(* IEC 61131-3 sources: daoli-st-library/DL_Process (part 22) *)

(* ---- FB_DL_BatteryTestCycler.st ---- *)
//==============================================================================
// 功能块：FB_DL_BatteryTestCycler ｜ 中文名称：单通道电池充放电工步机
// 所属子库：DL_Process ｜ 版本：v1.0.1 ｜ 兼容：CODESYS V3.5+ / TwinCAT 3 / 汇川 InoProShop
// 功能描述：单体电芯充放电测试工步机：静置 → 恒流充电 → 恒压充电 → 静置 → 恒流放电 →
//           静置 → 完成，逐工步按终止判据切相；充/放电容量按安时积分统计（LREAL 累加
//           防精度损失）；温度与电压安全域逐拍硬判，越限当拍断流并进故障相（锂电热失控
//           不可逆，安全路径优先级最高）。工步超时按「本工步独立计时」判定，禁跨相累计。
//           本件是单通道工步机：不调度多通道、不做通道仲裁与分配（多通道调度归
//           序号 19 的 FormationsChannelMgr），对外只以电流设定 / 电压限值与工步状态
//           布尔快照交互，两件互不包含。
// 开源溯源 (Origin)：道莅原创实现（参考 公开工程惯例 分类与参数域）
// 单位表：电压[V] / 电流[A]（放电为负）/ 温度[摄氏度] / 静置时长[min] / 工步超时[min] /
//         容量[Ah] / 容量比[百分数] / 扫描间隔[ms] / 工步已历时[ms] / 样本数[拍]
// 错误码表：16#0005_0406 信息级（工步切相提示，含「因终止判据达成而提前切相」与静置
//           到时，不置 bError）/ 16#0005_0407 信息级（容量统计饱和触顶，不置 bError）/
//           16#0005_034B 故障级（温度越上限或电压越安全域，或安全判据量（温度/电压/
//           电流）非有限——非有限按越限处置，强制断流，置 bError）/ 16#0005_034C 故障级
//           （单工步超时，工艺卡死，置 bError + 断流）/ 16#0005_034D 故障级（组态非法：
//           额定容量/电流设定/电压域/超时非正或非有限，以及状态机 ELSE 非法状态兜底）。
//           034D 的共用反证句：组态非法与非法状态在现有输出组合下不可观测出差异（均为
//           bError + fCurrentSetA = 0 + eStep 不推进 + bValid 撤），§3 未给本件独立组态槽，
//           故显式复用不越段。
// 状态机：E_DL_BatteryCycleState（eIdle=0 待机 / eRestInit=10 充电前静置 / eCcCharge=20
//           恒流充电 / eCvCharge=30 恒压充电 / eRestMid=40 放前静置 / eDiscCharge=50 恒流
//           放电 / eRestFinal=60 放后静置 / eDone=70 完成 / eFault=99 故障兜底），CASE 含
//           ELSE 兜底，ELSE 置 034D 且断流、eStep 回 eIdle。
// 边界行为：① 安全侧优先：温度 > fTempMaxC 或电压越 [fVoltMinV, fVoltMaxV] → 故障 034B
//           + fCurrentSetA := 0.0 + 进 eFault（每拍先判安全判据，先于任何工步推进）；
//           ② 单工步超 tMaxStep → 故障 034C，工步计时器在每次切相时清零（禁相内累计，
//           R40 家族）；③ 额定容量/电流/电压域/超时组态非法 → 034D 组态分支（映射见
//           错误码表反证句）；④ 容量积分 Ah += |I| x Δt/3600，LREAL 累加并饱和；⑤ CV
//           终止：|I| < fCutoffCurrentA 连续 nCvHoldSamples 拍才切相（防单点抖动误切）；
//           ⑥ bStop → 当拍 fCurrentSetA := 0 并回 eIdle（不等待工步收尾）；⑦ 失能走同一
//           安全侧路径（fCurrentSetA := 0）。bStart 取上升沿，bStepDone 为单拍脉冲。
// 修订历史：v1.0.0 2026-11-17 首版（R25 派单 · §4.15）
//           v1.0.1 2026-11-17 终审补 eFault 独立 CASE 标签（对外引脚契约零变更）：原实现 eFault(99)
//           无标签，落进 ELSE 兜底支路每拍把真因码 034B/034C 覆盖成 034D「非法状态」，激励消失后
//           诊断失真（故障仍锁存、安全侧不变，属诊断保真度缺陷）。同批另有 6 件存在同类标签缺失
//           （ParticleCounterStat / CoolingTowerApproachCalc / InverterGridSync / HeatPumpDefrost /
//           DuctStaticReset / DewpointReset），已按 R106 第二档挂账下轮统一修并加机检规则。
//==============================================================================
(*------------------------------------------------------------------------------
 * 枚举: E_DL_BatteryCycleState（归属 DL_Process，与 FB_DL_BatteryTestCycler 同文件）
 *       工步号与 §4.15 顺序一一对应；数值步长留空位便于插工步
 *----------------------------------------------------------------------------*)
TYPE E_DL_BatteryCycleState :
(
    eIdle       := 0,   // 待机：电流设定 0，等待 bStart / Idle, current setpoint 0, waiting for start
    eRestInit   := 10,  // 充电前静置：时长 tRestCharge / Pre-charge rest, duration tRestCharge
    eCcCharge   := 20,  // 恒流充电：电流 = fCcCurrentA，终止判据 电压达 fCvVoltV / Constant-current charge
    eCvCharge   := 30,  // 恒压充电：电压限 = fCvVoltV，终止判据 电流降至 fCutoffCurrentA / Constant-voltage charge
    eRestMid    := 40,  // 放前静置：时长 tRestCharge / Pre-discharge rest, duration tRestCharge
    eDiscCharge := 50,  // 恒流放电：电流 = -fDiscCurrentA，终止判据 电压降至 fDiscCutoffV / Constant-current discharge
    eRestFinal  := 60,  // 放后静置：时长 tRestDisc / Post-discharge rest, duration tRestDisc
    eDone       := 70,  // 完成：电流设定 0，容量统计保持 / Done, current 0, capacity statistics held
    eFault      := 99   // 故障兜底：越限/超时/组态非法/非法状态 / Fault fallback
);
END_TYPE

(*==============================================================================
 * 功能块: FB_DL_BatteryTestCycler
 * 调用约定: 每个扫描周期无条件调用一次；uDeltaTimeMs 必须注入真实任务间隔。
 *============================================================================*)
FUNCTION_BLOCK FB_DL_BatteryTestCycler
VAR_INPUT
    fVoltV          : LREAL;                       // 实测电压 [V] / Measured voltage [V]
    fCurrentA       : LREAL;                       // 实测电流 [A]，放电为负 / Measured current [A], negative while discharging
    fTempC          : LREAL;                       // 实测温度 [摄氏度] / Measured temperature [degC]
    fCcCurrentA     : LREAL;                       // 恒流充电电流设定 [A]，须 > 0 / Constant-current charge setpoint [A], must be > 0
    fCvVoltV        : LREAL;                       // 恒压充电电压点 [V] / Constant-voltage charge point [V]
    fCutoffCurrentA : LREAL;                       // 恒压段终止电流 [A]，须 >= 0 / CV termination current [A], must be >= 0
    fDiscCurrentA   : LREAL;                       // 放电电流设定 [A]，须 > 0（本件按负值下发）/ Discharge current setpoint [A], must be > 0, issued negative
    fDiscCutoffV    : LREAL;                       // 放电终止电压 [V] / Discharge termination voltage [V]
    tRestCharge     : TIME := T#10M;               // 充/放前静置时长 [min] / Pre-step rest duration [min]
    tRestDisc       : TIME := T#10M;               // 放后静置时长 [min] / Post-discharge rest duration [min]
    tMaxStep        : TIME := T#120M;              // 单工步超时 [min]，各工步独立计时 / Per-step timeout [min], timed per step
    fCapNomAh       : LREAL;                       // 额定容量 [Ah]，须 > 0（容量比分母）/ Rated capacity [Ah], must be > 0
    fVoltMaxV       : LREAL;                       // 安全域电压上限 [V] / Safety voltage ceiling [V]
    fVoltMinV       : LREAL;                       // 安全域电压下限 [V] / Safety voltage floor [V]
    fTempMaxC       : LREAL;                       // 温度上限 [摄氏度] / Temperature ceiling [degC]
    bStart          : BOOL;                        // 启动（取上升沿）/ Start, rising edge
    bStop           : BOOL;                        // 停止（电平，当拍断流）/ Stop, level, current dropped this scan
    bReset          : BOOL;                        // 复位，上升沿清故障与容量统计 / Reset, rising edge clears the fault and capacity statistics
    uDeltaTimeMs    : UDINT;                       // 扫描间隔 [ms]，调用方注入，禁系统时间函数 / Scan interval [ms], caller-injected
END_VAR
VAR_OUTPUT
    eStep           : E_DL_BatteryCycleState;      // 当前工步 / Current step
    fCurrentSetA    : LREAL;                       // 电流设定 [A]，故障拍立即 0 / Current setpoint [A], forced to 0 on any fault scan
    fVoltLimitV     : LREAL;                       // 电压限 [V]，随工步切换 / Voltage limit [V], follows the step
    fChargedAh      : LREAL;                       // 累计充电容量 [Ah]，饱和 / Accumulated charge capacity [Ah], saturating
    fDischargedAh   : LREAL;                       // 累计放电容量 [Ah]，饱和 / Accumulated discharge capacity [Ah], saturating
    fCapacityRatioPct : LREAL;                     // 容量比 [百分数] = 放电 Ah / 额定 Ah x 100 / Capacity ratio [percent]
    bStepDone       : BOOL;                        // 工步完成单拍脉冲（切相当拍 TRUE）/ Single-scan step-done pulse
    tStepElapsed    : TIME;                        // 本工步已历时 [ms] / Elapsed time of the current step [ms]
    eErr            : UDINT;                       // 错误码，0 = 无错，码位 16#0005_0406 起信息级、16#0005_034B 起故障级（分带见错误码表） / Error code, 0 = no error, band info/fault per the code table
    bError          : BOOL;                        // 故障级标志，仅故障级错误置位 / Fault-class flag, set only on fault-level codes
    bValid          : BOOL;                        // 工步输出可用标志，失能/故障闸显式 FALSE / Step outputs usable flag, explicit FALSE on disable/fault gates
END_VAR
VAR
    fbReset         : R_TRIG;                      // 复位上升沿检测实例 / Reset rising edge detector
    fbStart         : R_TRIG;                      // 启动上升沿检测实例 / Start rising edge detector
    uStepMs         : UDINT;                       // 本工步累计历时 [ms]，切相即清零 / Elapsed time of this step [ms], cleared on every transition
    uDtEff          : UDINT;                       // 钳位后的扫描间隔 [ms] / Clamped scan interval [ms]
    uMaxStepMs      : UDINT;                       // 工步超时门限 [ms] / Step timeout threshold [ms]
    uRestChgMs      : UDINT;                       // 充/放前静置门限 [ms] / Pre-step rest threshold [ms]
    uRestDiscMs     : UDINT;                       // 放后静置门限 [ms] / Post-discharge rest threshold [ms]
    fDtH            : LREAL;                       // 扫描间隔换算成小时 [h] / Scan interval in hours [h]
    fAbsCurrentA    : LREAL;                       // 实测电流绝对值 [A] / Absolute measured current [A]
    fAhStep         : LREAL;                       // 本拍容量增量 [Ah] / Capacity increment of this scan [Ah]
    nCvHoldCnt      : INT;                         // CV 终止判据连续满足拍数 [拍] / Consecutive CV-cutoff samples [scans]
    bCapSat         : BOOL;                        // 容量积分饱和标志 / Capacity saturation flag
    bStepChanged    : BOOL;                        // 本拍发生切相标志 / Step changed this scan
    bRestChgDone    : BOOL;                        // 静置到时（用充电侧时长）/ Rest elapsed with the charge-side duration
    bRestDiscDone   : BOOL;                        // 静置到时（用放电侧时长）/ Rest elapsed with the discharge-side duration
    bCvCutoff       : BOOL;                        // CV 终止判据满足 / CV termination criterion satisfied
    bDiscCutoff     : BOOL;                        // 放电终止判据满足 / Discharge termination criterion satisfied
    bCcReached      : BOOL;                        // CC 段电压已达 CV 点 / CC reached the CV point
    bNonFinSafe     : BOOL;                        // 安全判据量非有限标志 / Safety-class non-finite flag
    bNonFinCfg      : BOOL;                        // 组态量非有限标志 / Configuration non-finite flag
    bFirstScan      : BOOL := TRUE;                // 上电首拍标志 / First-scan flag
END_VAR
VAR CONSTANT
    DL_BTC_CODE_INFO_1 : UDINT := 16#0005_0406;    // 信息级槽 1（工步切相提示） / info slot 1
    DL_BTC_CODE_INFO_2 : UDINT := 16#0005_0407;    // 信息级槽 2（容量统计饱和） / info slot 2
    DL_BTC_CODE_FLT_1  : UDINT := 16#0005_034B;    // 故障级槽 1（温度/电压越限，强制断流） / fault slot 1
    DL_BTC_CODE_FLT_2  : UDINT := 16#0005_034C;    // 故障级槽 2（工步超时，工艺卡死） / fault slot 2
    DL_BTC_CODE_FLT_3  : UDINT := 16#0005_034D;    // 故障级槽 3（组态非法/非法状态兜底） / fault slot 3
    DL_BTC_CV_HOLD     : INT := 5;                 // CV 终止判据连续确认拍数 [拍] / CV cutoff confirmation samples [scans]
    DL_BTC_AH_MAX      : LREAL := 100000.0;        // 容量积分饱和上限 [Ah] / Capacity saturation ceiling [Ah]
    DL_BTC_DT_MIN_MS   : UDINT := 1;               // 扫描间隔下限 [ms]，防除零与死判 / Scan interval floor [ms]
    DL_BTC_SEC_PER_H   : LREAL := 3600.0;          // 秒转小时系数 [s/h] / Seconds per hour
    DL_BTC_MS_PER_S    : LREAL := 1000.0;          // 毫秒转秒系数 [ms/s] / Milliseconds per second
    DL_BTC_PCT         : LREAL := 100.0;           // 百分数系数 [百分数] / Percent factor
    DL_BTC_ZERO        : LREAL := 0.0;             // 零值常量，避免裸字面量 [—] / Zero constant, avoids a bare literal
    DL_BTC_TOL         : LREAL := 1.0E-6;          // 浮点比较容差 [—] / Float comparison tolerance
    DL_BTC_INF         : LREAL := 1.7976931348623157E308; // LREAL 幅值上限，Inf 判据 / LREAL magnitude ceiling
END_VAR

(*------------------------------------------------------------------------------
 * 段 1｜无条件刷新区（红线 5）：复位/启动沿检测在任何分支之外周期调用；
 *       bStepDone 为单拍脉冲，逐拍先清（调用方读到的仍是本拍值）
 *----------------------------------------------------------------------------*)
bStepDone := FALSE;                                // 单拍脉冲先清（自清机制）/ single-scan pulse cleared first
fCurrentSetA := DL_BTC_ZERO;                       // 电流设定默认 0：任何未显式赋值的路径都断流 / default 0, any unassigned path is de-energised
fVoltLimitV := DL_BTC_ZERO;                        // 电压限默认 0 / voltage limit defaults to zero
fbReset(CLK := bReset);                            // 复位沿检测无条件刷新 / reset edge refreshed unconditionally
fbStart(CLK := bStart);                            // 启动沿检测无条件刷新 / start edge refreshed unconditionally

(*------------------------------------------------------------------------------
 * 段 2｜复位沿处理（改写置于沿后，防吞沿 R39）：清故障与容量统计
 *----------------------------------------------------------------------------*)
IF fbReset.Q THEN
    eStep := E_DL_BatteryCycleState.eIdle;
    eErr   := 16#0000_0000;                        // 复位清码 / reset clears the code
    bError := FALSE;                               // 复位清故障 / reset clears the fault
    fChargedAh := DL_BTC_ZERO;                     // 充电容量清 / charge capacity cleared
    fDischargedAh := DL_BTC_ZERO;                  // 放电容量清 / discharge capacity cleared
    fCapacityRatioPct := DL_BTC_ZERO;              // 容量比清 / capacity ratio cleared
    uStepMs := 16#0000_0000;                       // 工步计时清 / step timer cleared
    nCvHoldCnt := 0;                               // CV 确认计数清 / CV hold counter cleared
    bCapSat := FALSE;                              // 饱和标志清 / saturation flag cleared
    bFirstScan := TRUE;                            // 重新首拍化 / re-initialize first scan
END_IF

(*------------------------------------------------------------------------------
 * 段 3｜非有限输入闸：安全判据量（温度/电压/电流）非有限 → 按越限处置（034B，断流）；
 *       组态量非有限 → 034D 组态分支。分两类是因为前者的正确处置是「当拍断流」，
 *       后者是「拒绝启动」
 *----------------------------------------------------------------------------*)
bNonFinSafe := (fVoltV <> fVoltV) OR (ABS(fVoltV) >= DL_BTC_INF)
            OR (fCurrentA <> fCurrentA) OR (ABS(fCurrentA) >= DL_BTC_INF)
            OR (fTempC <> fTempC) OR (ABS(fTempC) >= DL_BTC_INF);   // 安全判据量非有限 / safety-class non-finite
bNonFinCfg := (fCcCurrentA <> fCcCurrentA) OR (ABS(fCcCurrentA) >= DL_BTC_INF)
           OR (fCvVoltV <> fCvVoltV) OR (ABS(fCvVoltV) >= DL_BTC_INF)
           OR (fCutoffCurrentA <> fCutoffCurrentA) OR (ABS(fCutoffCurrentA) >= DL_BTC_INF)
           OR (fDiscCurrentA <> fDiscCurrentA) OR (ABS(fDiscCurrentA) >= DL_BTC_INF)
           OR (fDiscCutoffV <> fDiscCutoffV) OR (ABS(fDiscCutoffV) >= DL_BTC_INF)
           OR (fCapNomAh <> fCapNomAh) OR (ABS(fCapNomAh) >= DL_BTC_INF)
           OR (fVoltMaxV <> fVoltMaxV) OR (ABS(fVoltMaxV) >= DL_BTC_INF)
           OR (fVoltMinV <> fVoltMinV) OR (ABS(fVoltMinV) >= DL_BTC_INF)
           OR (fTempMaxC <> fTempMaxC) OR (ABS(fTempMaxC) >= DL_BTC_INF);   // 组态量非有限 / configuration non-finite
IF bNonFinSafe THEN
    eStep := E_DL_BatteryCycleState.eFault;        // 进故障相 / enter fault state
    eErr   := DL_BTC_CODE_FLT_1;                   // 故障级：安全判据不可判，按越限处置 / fault: safety values undecidable, treated as out of range
    bError := TRUE;                                // 故障级必置 bError（R45 配对）/ fault-class pairs with bError
    fCurrentSetA := DL_BTC_ZERO;                   // 当拍断流（安全路径最高优先）/ current dropped this scan
    fVoltLimitV := DL_BTC_ZERO;                    // 电压限撤 / voltage limit dropped
    bValid := FALSE;                               // 故障闸显式不可用（R72）/ explicit FALSE on the fault gate
    RETURN;
END_IF
IF bNonFinCfg THEN
    eStep := E_DL_BatteryCycleState.eFault;        // 进故障相 / enter fault state
    eErr   := DL_BTC_CODE_FLT_3;                   // 故障级：组态非法（映射见错误码表）/ fault: invalid configuration, mapping per the code table
    bError := TRUE;                                // 故障级必置 bError（R45 配对）/ fault-class pairs with bError
    fCurrentSetA := DL_BTC_ZERO;                   // 断流 / current dropped
    fVoltLimitV := DL_BTC_ZERO;                    // 电压限撤 / voltage limit dropped
    bValid := FALSE;                               // 故障闸显式不可用（R72）/ explicit FALSE on the fault gate
    RETURN;
END_IF

(*------------------------------------------------------------------------------
 * 段 4｜组态域闸（034D 组态分支，先判后除：容量比分母在此被证明为正）
 *----------------------------------------------------------------------------*)
IF (fCapNomAh <= DL_BTC_TOL) OR (fVoltMaxV <= fVoltMinV + DL_BTC_TOL)
   OR (fCcCurrentA <= DL_BTC_TOL) OR (fDiscCurrentA <= DL_BTC_TOL)
   OR (fCutoffCurrentA < DL_BTC_ZERO)
   OR (DINT_TO_UDINT(TIME_TO_DINT(tMaxStep)) = 16#00000000) THEN
    eStep := E_DL_BatteryCycleState.eFault;        // 进故障相 / enter fault state
    eErr   := DL_BTC_CODE_FLT_3;                   // 故障级：组态非法 / fault: invalid configuration
    bError := TRUE;                                // 故障级必置 bError（R45 配对）/ fault-class pairs with bError
    fCurrentSetA := DL_BTC_ZERO;                   // 断流 / current dropped
    fVoltLimitV := DL_BTC_ZERO;                    // 电压限撤 / voltage limit dropped
    bValid := FALSE;                               // 故障闸显式不可用（R72）/ explicit FALSE on the fault gate
    RETURN;
END_IF

(*------------------------------------------------------------------------------
 * 段 5｜安全域硬判（最高优先，先于任何工步推进）：温度越上限或电压越安全域 →
 *       034B + 当拍断流 + 进故障相。故障锁存至 bReset（热失控不可逆）
 *----------------------------------------------------------------------------*)
IF (fTempC > fTempMaxC) OR (fVoltV > fVoltMaxV + DL_BTC_TOL) OR (fVoltV < fVoltMinV - DL_BTC_TOL) THEN
    eStep := E_DL_BatteryCycleState.eFault;        // 进故障相 / enter fault state
    eErr   := DL_BTC_CODE_FLT_1;                   // 故障级：温度/电压越限 / fault: temperature or voltage out of range
    bError := TRUE;                                // 故障级必置 bError（R45 配对）/ fault-class pairs with bError
    fCurrentSetA := DL_BTC_ZERO;                   // 当拍断流（安全侧）/ current dropped this scan, safe side
    fVoltLimitV := DL_BTC_ZERO;                    // 电压限撤 / voltage limit dropped
    bValid := FALSE;                               // 故障闸显式不可用（R72）/ explicit FALSE on the fault gate
    RETURN;
END_IF

(*------------------------------------------------------------------------------
 * 段 6｜工步计时：仅活动工步累计（切相清零），静置/完成/待机不累计
 *----------------------------------------------------------------------------*)
IF uDeltaTimeMs < DL_BTC_DT_MIN_MS THEN
    uDtEff := DL_BTC_DT_MIN_MS;                     // 间隔过小按下限，防死等 / floored interval prevents a dead wait
ELSE
    uDtEff := uDeltaTimeMs;                         // 间隔原值 / interval as-is
END_IF
IF (eStep <> E_DL_BatteryCycleState.eIdle) AND (eStep <> E_DL_BatteryCycleState.eDone)
   AND (eStep <> E_DL_BatteryCycleState.eFault) THEN
    IF uStepMs < 16#FFFF_FFFE THEN
        uStepMs := uStepMs + uDtEff;                // 本工步累计 [ms] / accumulate the current step [ms]
    END_IF
END_IF
uMaxStepMs := DINT_TO_UDINT(TIME_TO_DINT(tMaxStep));       // 超时门限 [ms] / timeout threshold [ms]
uRestChgMs := DINT_TO_UDINT(TIME_TO_DINT(tRestCharge));    // 充/放前静置门限 [ms] / pre-step rest threshold [ms]
uRestDiscMs := DINT_TO_UDINT(TIME_TO_DINT(tRestDisc));     // 放后静置门限 [ms] / post-discharge rest threshold [ms]

(*------------------------------------------------------------------------------
 * 段 7｜工步超时（034C）：各工步独立计时，切相即清零，禁相内累计（R40 家族）
 *----------------------------------------------------------------------------*)
IF (eStep <> E_DL_BatteryCycleState.eIdle) AND (eStep <> E_DL_BatteryCycleState.eDone)
   AND (eStep <> E_DL_BatteryCycleState.eFault) AND (uStepMs > uMaxStepMs) THEN
    eStep := E_DL_BatteryCycleState.eFault;        // 进故障相 / enter fault state
    eErr   := DL_BTC_CODE_FLT_2;                   // 故障级：工步超时，工艺卡死 / fault: step timeout, process stuck
    bError := TRUE;                                // 故障级必置 bError（R45 配对）/ fault-class pairs with bError
    fCurrentSetA := DL_BTC_ZERO;                   // 断流 / current dropped
    fVoltLimitV := DL_BTC_ZERO;                    // 电压限撤 / voltage limit dropped
    bValid := FALSE;                               // 故障闸显式不可用（R72）/ explicit FALSE on the fault gate
    RETURN;
END_IF

(*------------------------------------------------------------------------------
 * 段 8｜容量安时积分：Ah += |I| x Δt/3600（LREAL 累加防精度损失，饱和防溢出）
 *----------------------------------------------------------------------------*)
fDtH := UDINT_TO_LREAL(uDtEff) / DL_BTC_MS_PER_S / DL_BTC_SEC_PER_H;   // 间隔换算成小时 [h] / interval in hours
fAbsCurrentA := ABS(fCurrentA);                    // 电流绝对值 [A] / absolute current [A]
fAhStep := fAbsCurrentA * fDtH;                     // 本拍容量增量 [Ah] / capacity increment [Ah]
IF (eStep = E_DL_BatteryCycleState.eCcCharge) OR (eStep = E_DL_BatteryCycleState.eCvCharge) THEN
    IF fChargedAh < DL_BTC_AH_MAX THEN
        fChargedAh := fChargedAh + fAhStep;         // 充电容量累加 [Ah] / charge capacity accumulation
        IF fChargedAh >= DL_BTC_AH_MAX THEN
            fChargedAh := DL_BTC_AH_MAX;            // 饱和钳位 [Ah] / saturation clamp
            bCapSat := TRUE;                        // 饱和标志 / saturation flag
        END_IF
    ELSE
        bCapSat := TRUE;                            // 已在饱和点 / already saturated
    END_IF
END_IF
IF eStep = E_DL_BatteryCycleState.eDiscCharge THEN
    IF fDischargedAh < DL_BTC_AH_MAX THEN
        fDischargedAh := fDischargedAh + fAhStep;   // 放电容量累加 [Ah] / discharge capacity accumulation
        IF fDischargedAh >= DL_BTC_AH_MAX THEN
            fDischargedAh := DL_BTC_AH_MAX;         // 饱和钳位 [Ah] / saturation clamp
            bCapSat := TRUE;                        // 饱和标志 / saturation flag
        END_IF
    ELSE
        bCapSat := TRUE;                            // 已在饱和点 / already saturated
    END_IF
END_IF
fCapacityRatioPct := fDischargedAh / fCapNomAh * DL_BTC_PCT;   // 容量比（除子已由段 4 证明为正）[百分数] / capacity ratio, divisor proven positive
tStepElapsed := UDINT_TO_TIME(uStepMs);            // 本工步已历时 [ms] / elapsed time of the current step

(*------------------------------------------------------------------------------
 * 段 9｜停止闸（电平，当拍生效）：断流并回待机，不等待工步收尾（安全侧）
 *----------------------------------------------------------------------------*)
IF bStop THEN
    eStep := E_DL_BatteryCycleState.eIdle;         // 回待机 / back to idle
    fCurrentSetA := DL_BTC_ZERO;                   // 当拍断流 / current dropped this scan
    fVoltLimitV := DL_BTC_ZERO;                    // 电压限撤 / voltage limit dropped
    uStepMs := 16#0000_0000;                       // 工步计时清 / step timer cleared
    nCvHoldCnt := 0;                               // CV 确认计数清 / CV hold counter cleared
    eErr := 16#0000_0000;                          // 停止清信息码 / stop clears info codes
    bValid := FALSE;                               // 停止闸显式不可用（R72）/ explicit FALSE on the stop gate
    RETURN;
END_IF

(*------------------------------------------------------------------------------
 * 段 10｜工步状态机：CASE 含 ELSE 兜底（非法状态 → 034D + 断流 + 回待机）
 *       切相一律：uStepMs := 0（禁相内累计）+ bStepDone 单拍脉冲
 *----------------------------------------------------------------------------*)
bStepChanged := FALSE;                             // 切相标志逐拍重判 / transition flag re-judged per scan
bCcReached := (fVoltV >= fCvVoltV - DL_BTC_TOL);            // CC 段电压达 CV 点 / CC reached the CV point
bCvCutoff := (fAbsCurrentA < fCutoffCurrentA + DL_BTC_TOL);  // CV 终止判据 / CV termination predicate
bDiscCutoff := (fVoltV <= fDiscCutoffV + DL_BTC_TOL);        // 放电终止判据 / discharge termination predicate
bRestChgDone := (uStepMs >= uRestChgMs);           // 充/放前静置到时 / pre-step rest elapsed
bRestDiscDone := (uStepMs >= uRestDiscMs);         // 放后静置到时 / post-discharge rest elapsed
IF bCvCutoff THEN
    IF nCvHoldCnt < DL_BTC_CV_HOLD THEN
        nCvHoldCnt := nCvHoldCnt + 1;              // 连续满足拍数饱和自增 [拍] / saturating consecutive-sample counter
    END_IF
ELSE
    nCvHoldCnt := 0;                               // 判据断链即清零（防单点抖动误切）/ counter cleared on any drop-out
END_IF

CASE eStep OF

    E_DL_BatteryCycleState.eIdle:
        fCurrentSetA := DL_BTC_ZERO;               // 待机断流 / de-energised in idle
        fVoltLimitV := DL_BTC_ZERO;                // 待机无电压限 / no voltage limit in idle
        uStepMs := 16#0000_0000;                   // 待机不计时 / no timing in idle
        nCvHoldCnt := 0;                           // CV 计数清 / CV counter cleared
        eErr := 16#0000_0000;                      // 待机无错 / no error in idle
        bError := FALSE;                           // 待机无故障 / no fault in idle
        IF fbStart.Q THEN
            eStep := E_DL_BatteryCycleState.eRestInit;   // 上升沿启动：先进充电前静置 / start edge enters the pre-charge rest
            uStepMs := 16#0000_0000;               // 新工步计时清零 / new step timer cleared
            bStepChanged := TRUE;                  // 切相标志 / transition flag
            bFirstScan := FALSE;                   // 首拍标志清除 / first-scan flag cleared
        END_IF

    E_DL_BatteryCycleState.eRestInit:
        fCurrentSetA := DL_BTC_ZERO;               // 静置断流 / de-energised while resting
        fVoltLimitV := DL_BTC_ZERO;                // 静置无电压限 / no voltage limit while resting
        eErr := DL_BTC_CODE_INFO_1;                // 信息级：工步在静置相（切相提示）/ info: resting step
        bError := FALSE;                           // 信息级不置 bError / info never raises bError
        IF bRestChgDone THEN
            eStep := E_DL_BatteryCycleState.eCcCharge;   // 静置到时进恒流充电 / rest elapsed, enter CC charge
            uStepMs := 16#0000_0000;               // 新工步计时清零（禁相内累计）/ new step timer cleared
            bStepChanged := TRUE;                  // 切相标志 / transition flag
        END_IF

    E_DL_BatteryCycleState.eCcCharge:
        fCurrentSetA := fCcCurrentA;               // 恒流充电电流 [A] / CC charge current [A]
        fVoltLimitV := fVoltMaxV;                  // 电压限取安全域上限 [V] / voltage limit at the safety ceiling [V]
        eErr := DL_BTC_CODE_INFO_1;                // 信息级：工步在恒流充电相 / info: CC charge step
        bError := FALSE;                           // 信息级不置 bError / info never raises bError
        IF bCcReached THEN
            eStep := E_DL_BatteryCycleState.eCvCharge;   // 电压达 CV 点切恒压（终止判据达成）/ CV point reached, enter CV
            uStepMs := 16#0000_0000;               // 新工步计时清零 / new step timer cleared
            nCvHoldCnt := 0;                       // CV 计数复位 / CV counter reset
            bStepChanged := TRUE;                  // 切相标志 / transition flag
        END_IF

    E_DL_BatteryCycleState.eCvCharge:
        fCurrentSetA := fCcCurrentA;               // 恒压段电流上限仍为设定值 [A] / CV current ceiling stays at the setpoint [A]
        fVoltLimitV := fCvVoltV;                   // 恒压点 [V] / CV point [V]
        eErr := DL_BTC_CODE_INFO_1;                // 信息级：工步在恒压充电相 / info: CV charge step
        bError := FALSE;                           // 信息级不置 bError / info never raises bError
        IF nCvHoldCnt >= DL_BTC_CV_HOLD THEN
            eStep := E_DL_BatteryCycleState.eRestMid;    // 电流连续 5 拍低于终止值切静置 / cutoff sustained, enter the pre-discharge rest
            uStepMs := 16#0000_0000;               // 新工步计时清零 / new step timer cleared
            nCvHoldCnt := 0;                       // CV 计数复位 / CV counter reset
            bStepChanged := TRUE;                  // 切相标志 / transition flag
        END_IF

    E_DL_BatteryCycleState.eRestMid:
        fCurrentSetA := DL_BTC_ZERO;               // 静置断流 / de-energised while resting
        fVoltLimitV := DL_BTC_ZERO;                // 静置无电压限 / no voltage limit while resting
        eErr := DL_BTC_CODE_INFO_1;                // 信息级：工步在放前静置相 / info: pre-discharge rest step
        bError := FALSE;                           // 信息级不置 bError / info never raises bError
        IF bRestChgDone THEN
            eStep := E_DL_BatteryCycleState.eDiscCharge;   // 静置到时进恒流放电 / rest elapsed, enter CC discharge
            uStepMs := 16#0000_0000;               // 新工步计时清零 / new step timer cleared
            bStepChanged := TRUE;                  // 切相标志 / transition flag
        END_IF

    E_DL_BatteryCycleState.eDiscCharge:
        fCurrentSetA := -ABS(fDiscCurrentA);       // 放电电流按负值下发（放电为负）[A] / discharge issued negative [A]
        fVoltLimitV := fDiscCutoffV;               // 放电终止电压作为下限语义的限值 [V] / discharge cut-off as the limit [V]
        eErr := DL_BTC_CODE_INFO_1;                // 信息级：工步在恒流放电相 / info: CC discharge step
        bError := FALSE;                           // 信息级不置 bError / info never raises bError
        IF bDiscCutoff THEN
            eStep := E_DL_BatteryCycleState.eRestFinal;   // 电压达放电终止切静置 / cut-off reached, enter the final rest
            uStepMs := 16#0000_0000;               // 新工步计时清零 / new step timer cleared
            bStepChanged := TRUE;                  // 切相标志 / transition flag
        END_IF

    E_DL_BatteryCycleState.eRestFinal:
        fCurrentSetA := DL_BTC_ZERO;               // 静置断流 / de-energised while resting
        fVoltLimitV := DL_BTC_ZERO;                // 静置无电压限 / no voltage limit while resting
        eErr := DL_BTC_CODE_INFO_1;                // 信息级：工步在放后静置相 / info: post-discharge rest step
        bError := FALSE;                           // 信息级不置 bError / info never raises bError
        IF bRestDiscDone THEN
            eStep := E_DL_BatteryCycleState.eDone; // 放后静置到时转完成 / post-discharge rest elapsed, done
            uStepMs := 16#0000_0000;               // 新工步计时清零 / new step timer cleared
            bStepChanged := TRUE;                  // 切相标志 / transition flag
        END_IF

    E_DL_BatteryCycleState.eDone:
        fCurrentSetA := DL_BTC_ZERO;               // 完成态断流 / de-energised when done
        fVoltLimitV := DL_BTC_ZERO;                // 完成态无电压限 / no voltage limit when done
        eErr := 16#0000_0000;                      // 完成无错 / no error when done
        bError := FALSE;                           // 完成无故障 / no fault when done
        IF fbStart.Q THEN
            eStep := E_DL_BatteryCycleState.eRestInit;   // 再次启动重跑一轮 / a new start edge runs another cycle
            uStepMs := 16#0000_0000;               // 计时清零 / timer cleared
            fChargedAh := DL_BTC_ZERO;             // 容量统计重新起算 / capacity statistics restart
            fDischargedAh := DL_BTC_ZERO;          // 容量统计重新起算 / capacity statistics restart
            bStepChanged := TRUE;                  // 切相标志 / transition flag
        END_IF

    E_DL_BatteryCycleState.eFault:
        // v1.0.1 修正：eFault 是合法故障态，必须有独立 CASE 标签。原实现缺此标签，eFault(99) 每拍落进
        // ELSE 兜底支路，把段 3/4/5/7 已判定的 034B（越限断流）/034C（工步超时）覆盖成 034D（非法状态），
        // 激励消失（温度回到域内、超时条件不再成立）后真因码即丢失，诊断只能看到「非法状态」。
        // 本相只做安全侧输出与故障码保持，故障码改写一律归入口闸，零码兜底由段 11 统一处理。
        fCurrentSetA := DL_BTC_ZERO;               // 故障相断流（安全值而非上次值）/ zeroed in fault, never the last value
        fVoltLimitV := DL_BTC_ZERO;                // 电压限撤 / voltage limit dropped
        bError := TRUE;                            // 故障级必置 bError（R45 配对）/ fault-class pairs with bError
        // eErr 保持：不得在本相改写（禁 034B/034C → 034D 覆盖）

    ELSE
        eStep := E_DL_BatteryCycleState.eFault;    // 非法状态兜底 / illegal-state fallback
        eErr := DL_BTC_CODE_FLT_3;                 // 故障级兜底：非法状态 / fault fallback: illegal state
        bError := TRUE;                            // 故障级必置 bError（R45 配对）/ fault-class pairs with bError
        fCurrentSetA := DL_BTC_ZERO;               // 断流安全侧 / current dropped, safe side
        fVoltLimitV := DL_BTC_ZERO;                // 电压限撤 / voltage limit dropped

END_CASE

(*------------------------------------------------------------------------------
 * 段 11｜故障相最终闸与出口收口：故障态一律断流（安全值而非上次值），
 *       切相脉冲与饱和提示在本拍出口统一落定
 *----------------------------------------------------------------------------*)
IF eStep = E_DL_BatteryCycleState.eFault THEN
    fCurrentSetA := DL_BTC_ZERO;                   // 故障拍立即 0（安全侧，不保留上次设定）/ zero on any fault scan, never the last value
    fVoltLimitV := DL_BTC_ZERO;                    // 电压限撤 / voltage limit dropped
    bError := TRUE;                                // 故障级必置 bError（R45 配对）/ fault-class pairs with bError
    IF eErr = 16#0000_0000 THEN
        eErr := DL_BTC_CODE_FLT_3;                 // 入口无码时按非法状态兜底（R45：bError 必须有对应码）/ illegal-state fallback
    END_IF
    IF bReset THEN
        eStep := E_DL_BatteryCycleState.eIdle;     // 仅复位可退出故障相（热失控类故障不得自愈）/ only reset leaves the fault state
    END_IF
ELSE
    IF bCapSat THEN
        eErr := DL_BTC_CODE_INFO_2;                // 信息级：容量统计饱和（优先于切相提示）/ info: capacity saturation outranks the step hint
    END_IF
    IF bStepChanged THEN
        bStepDone := TRUE;                         // 切相当拍输出单拍脉冲 / single-scan pulse on a transition
        IF NOT bCapSat THEN
            eErr := DL_BTC_CODE_INFO_1;            // 信息级：工步切相提示 / info: step transition hint
        END_IF
    END_IF
END_IF
bValid := (eStep <> E_DL_BatteryCycleState.eFault);   // 许可类输出显式落定（R72）/ permission settled explicitly
END_FUNCTION_BLOCK

(* ---- FB_DL_BeltHeatRecovery.st ---- *)
(*
  ==================================================================
  组件名 Component  : FB_DL_BeltHeatRecovery
  分类   Category   : DL_Process
  版本   Version    : 1.0.0
  功能   Purpose    : 转轮热回收与输送联锁。按「转轮先启、输送后行、停输后吹扫」
                      的时序编排输送允许信号：转轮运行命令与反馈、过滤网状态、
                      火警联锁、防霜限温四条判据共同决定输送允许；停输后转轮
                      继续运行 tStopDelay 完成吹扫再停。同时按进排风温差算热回收
                      效率并给出效率达标标志。
  溯源   Origin     : 转轮热回收联锁为通用暖通时序语义；本件为 clean-room 实现，
                      仅借鉴来源分类与参数域组织（来源标签 roadmap-p2-hvac），
                      道莅原创设计，未复制任何闭源代码行。
  平台   Platform   : 纯 IEC 61131-3（TON / R_TRIG / REAL 运算，无私有库）
  作者   Author     : 道莅代码库 · PLC 编程专家（R55）
  ------------------------------------------------------------------
  同拍双窗配比约束（R100）：tStopDelay 必须大于等于 tStartDelay，保证吹扫窗
                      不短于启动窗；两窗职责分离：启动窗等转轮反馈，吹扫窗保
                      转轮续转，任一窗不得兼作另一窗用途。
  边界 Boundary     :
                      一 本件只出输送允许与转轮命令，不直接驱动风机变频器（属主边界）；
                      二 火警联锁优先级最高：撤转轮命令 + 撤输送允许 + 锁存至复位沿；
                      三 防霜判据成立时撤输送允许但保留转轮运行（防冻需转轮换热）；
                      四 过滤网异常撤输送允许但保留转轮运行（降级运行并置成因）；
                      五 无全局变量、无外部变量声明、无物理地址寻址。
  输出契约 Output contract:
                      bConvPermit 仅在运行相且转轮反馈到位、无火警、过滤网正常、
                      未触发防霜时为真（挂状态量，非单拍标志）；
                      fEffPct 在进排风温差不足 fMinDeltaTC 时保持上拍值并置 bEffOk 为假；
                      eCause 故障级成因与 bError 配对（R45），信息级永不置 bError。
  修订记录 Revision  :
    2026-11-20  v1.0.0  R55 首版（批 3 · 序号 14）
  ==================================================================
*)

TYPE E_DL_BhrState :
(
    eIdle      := 0,    // 空闲：转轮停、输送禁行 / idle, the wheel is stopped and the conveyor is inhibited
    eStartWait := 10,   // 启动等反馈：等转轮运行反馈与启动延时 / waiting for the wheel feedback and the start delay
    eRun       := 20,   // 运行：输送允许 / running, the conveyor is permitted
    ePurge     := 30,   // 吹扫：停输后转轮续转 / purge, the wheel keeps running after the conveyor stops
    eFault     := 90    // 故障：火警或组态非法锁存 / fault, fire alarm or illegal configuration latched
);
END_TYPE

TYPE E_DL_BhrCause :
(
    eNone       := 0,   // 无成因 / no cause
    eCfgIllegal := 1,   // 组态非法：时间窗配比反置或阈值越域（故障级，与 bError 配对）/ illegal config, window ratio inverted or a threshold out of domain
    eFireAlarm  := 2,   // 火警联锁动作（故障级，与 bError 配对，锁存至复位沿）/ fire alarm interlock tripped, a fault latched until the reset edge
    eFrost      := 3,   // 防霜动作，撤输送允许（信息级）/ frost protection tripped and the conveyor was inhibited, informational
    eFilterBad  := 4,   // 过滤网异常，撤输送允许（信息级）/ filter fault inhibited the conveyor, informational
    eNoWheelFb  := 5,   // 转轮反馈缺失，输送不放开（信息级）/ the wheel feedback is missing so the conveyor stays inhibited, informational
    eEffInvalid := 6    // 进排风温差不足，效率不更新（信息级）/ the temperature difference is too small and the efficiency holds, informational
);
END_TYPE

FUNCTION_BLOCK FB_DL_BeltHeatRecovery
VAR_INPUT
    bEnable      : BOOL := TRUE;             // 使能，失能时全部命令撤除 [-] / enable, all commands are withdrawn when disabled
    bReset       : BOOL := FALSE;           // 复位上升沿清故障锁存（火警须已消失）/ reset rising edge clears the fault latch, the fire alarm must be cleared first
    bConvRunCmd  : BOOL := FALSE;            // 输送运行请求（电平）[-] / conveyor run request, a level
    bWheelRunFb  : BOOL := FALSE;            // 转轮运行反馈 [-] / wheel running feedback
    bFilterOk    : BOOL := FALSE;            // 过滤网正常 [-] / filter healthy
    bFireAlarm   : BOOL := FALSE;            // 火警联锁源 [-] / fire alarm interlock source
    fExhaustC    : REAL := 20.0;             // 排风温度 [摄氏度] / exhaust air temperature [degree Celsius]
    fSupplyC     : REAL := 20.0;             // 送风温度（转轮后）[摄氏度] / supply air temperature after the wheel [degree Celsius]
    fFreshC      : REAL := 10.0;             // 新风温度（转轮前）[摄氏度] / fresh air temperature before the wheel [degree Celsius]
    fFrostLimitC : REAL := -5.0;             // 防霜限温 [摄氏度]，域 -60..10 / frost protection limit [degree Celsius], domain minus sixty to ten
    fMinDeltaTC  : REAL := 5.0;              // 效率计算的进排风最小温差 [开尔文]，域 大于零 / minimum exhaust to fresh difference for the efficiency calculation [Kelvin], domain above zero
    fEffMinPct   : REAL := 50.0;             // 效率达标阈 [百分比]，域 0..100 / efficiency pass threshold [percent], domain 0 to 100
    tStartDelay  : TIME := T#5S;             // 启动延时（转轮先启）[毫秒] / start delay so the wheel leads [millisecond]
    tStopDelay   : TIME := T#30S;            // 吹扫延时（输送后停）[毫秒]，须不短于启动延时 / purge delay so the wheel lags [millisecond], not shorter than the start delay
END_VAR
VAR_OUTPUT
    bConvPermit  : BOOL := FALSE;            // 输送允许 [-] / conveyor permit
    bWheelRunCmd : BOOL := FALSE;            // 转轮运行命令 [-] / wheel run command
    bFrostProtect: BOOL := FALSE;            // 防霜动作中 [-] / frost protection active
    bWheelFbOk   : BOOL := FALSE;            // 转轮反馈到位 [-] / wheel feedback present
    fEffPct      : REAL := 0.0;              // 热回收效率（锁存值）[百分比] / heat recovery efficiency, latched [percent]
    bEffOk       : BOOL := FALSE;            // 效率达标且本拍有效 [-] / efficiency passes and this scan is valid
    eState       : E_DL_BhrState := E_DL_BhrState.eIdle; // 相位出口 [枚举] / phase outlet [enum]
    eCause       : E_DL_BhrCause := E_DL_BhrCause.eNone; // 成因出口 [枚举] / cause outlet [enum]
    bError       : BOOL := FALSE;            // 故障锁存标志 [-] / fault latch flag
END_VAR
VAR
    rtReset      : R_TRIG;                   // 复位沿检测，段 0 无条件刷新 / reset edge detector, refreshed unconditionally in segment zero
    tonStart     : TON;                      // 启动延时，段 0 无条件刷新 / start delay, refreshed unconditionally in segment zero
    tonStop      : TON;                      // 吹扫延时，段 0 无条件刷新 / purge delay, refreshed unconditionally in segment zero
    _eState      : E_DL_BhrState := E_DL_BhrState.eIdle;  // 内部相位，CASE 唯一写入目标 / internal phase, the only CASE write target
    _eCause      : E_DL_BhrCause := E_DL_BhrCause.eNone;  // 信息级成因，每拍重算 / informational cause, recomputed every scan
    _eFaultCause : E_DL_BhrCause := E_DL_BhrCause.eNone;  // 故障级成因，锁存至复位沿 / fault cause, latched until the reset edge
    _bFault      : BOOL := FALSE;            // 故障锁存位 [-] / fault latch bit
    _bInit       : BOOL := FALSE;            // 首扫初始化完成标志（R310）/ first scan initialisation flag
    _bCfgBad     : BOOL := FALSE;            // 组态非法判定 [-] / illegal configuration verdict
    _bTempOk     : BOOL := FALSE;            // 三项温度均有限 [-] / all three temperatures finite
    _bEffBaseOk  : BOOL := FALSE;            // 效率分母可用 [-] / the efficiency denominator is usable
    _bFrost      : BOOL := FALSE;            // 防霜动作判定 [-] / frost protection verdict
    _bWheelFbOk  : BOOL := FALSE;            // 转轮反馈到位判定 [-] / wheel feedback verdict
    _bConvPermit : BOOL := FALSE;            // 输送允许判定 [-] / conveyor permit verdict
    _fEff         : REAL := 0.0;             // 效率工作值 [百分比] / efficiency working value [percent]
    _fEffHold     : REAL := 0.0;             // 效率保持块 [百分比] / efficiency holder [percent]
    _fDeltaT      : REAL := 0.0;             // 进排风温差（分母）[开尔文] / exhaust to fresh difference, the denominator [Kelvin]
    _fNum         : REAL := 0.0;             // 效率分子（送风减新风）[开尔文] / numerator, supply minus fresh [Kelvin]
END_VAR
VAR CONSTANT
    DL_BHR_EFF_MIN   : REAL := -100.0;       // 效率下限（负效率可能：转轮反向传热）[百分比] / efficiency floor, a negative value is possible [percent]
    DL_BHR_EFF_MAX   : REAL := 150.0;        // 效率上限 [百分比] / efficiency ceiling [percent]
    DL_BHR_FROST_MIN : REAL := -60.0;        // 防霜限温下限 [摄氏度] / frost limit floor [degree Celsius]
    DL_BHR_FROST_MAX : REAL := 10.0;         // 防霜限温上限 [摄氏度] / frost limit ceiling [degree Celsius]
    DL_BHR_DELTA_MAX : REAL := 200.0;        // 最小温差上限 [开尔文] / minimum difference ceiling [Kelvin]
    DL_BHR_TEMP_MAX  : REAL := 200.0;        // 温度量级上限（绝对值）[摄氏度] / temperature magnitude ceiling as an absolute value [degree Celsius]
END_VAR

// 段 0｜定时器与沿检测无条件周期刷新（禁入分支），IN 只串状态闸与业务闸 / segment 0, unconditional refresh with state and process gates on IN only
rtReset(CLK := bReset); // 复位沿无条件刷新 / unconditional refresh of the reset edge
tonStart(IN := (_eState = E_DL_BhrState.eStartWait) AND (NOT _bFault), PT := tStartDelay); // 启动延时，仅在等反馈相计时 / start delay timing only in the waiting phase
tonStop(IN := (_eState = E_DL_BhrState.ePurge) AND (NOT _bFault), PT := tStopDelay); // 吹扫延时，仅在吹扫相计时 / purge delay timing only in the purge phase

// 段 1｜首扫初始化（R310）/ segment 1, first scan initialisation
IF NOT _bInit THEN // 首扫一拍 / the very first scan
    _bInit := TRUE; // 置首扫完成标志 / raise the first scan flag
    _eState := E_DL_BhrState.eIdle; // 相位从空闲起步 / the phase starts from idle
    _eCause := E_DL_BhrCause.eNone; // 信息级成因清零 / clear the informational cause
    _eFaultCause := E_DL_BhrCause.eNone; // 故障级成因清零 / clear the fault cause
    _bFault := FALSE; // 故障锁存清零 / clear the fault latch
    _fEffHold := 0.0; // 效率保持块清零 / clear the efficiency holder
END_IF

// 段 2｜复位沿作用域：清故障锁存（火警必须已消失才允许解除，R152 可达性）/ segment 2, reset edge scope with a reachable release condition
IF rtReset.Q AND (NOT bFireAlarm) THEN // 复位沿且火警已消失 / reset edge with the fire alarm cleared
    _bFault := FALSE; // 作用域一：清故障锁存 / scope one, clear the fault latch
    _eFaultCause := E_DL_BhrCause.eNone; // 作用域一：清故障级成因 / scope one, clear the fault cause
    _eState := E_DL_BhrState.eIdle; // 作用域二：迁回空闲相 / scope two, migrate back to idle
END_IF

// 段 3｜组态域闸（R151 全覆盖）：双窗配比（R100）+ 阈值域 / segment 3, configuration domain gate including the window ratio
_bCfgBad := FALSE; // 组态非法预置假 / preset the illegal configuration verdict to false
IF tStopDelay < tStartDelay THEN // 吹扫窗短于启动窗，违反配比约束 / the purge window is shorter than the start window
    _bCfgBad := TRUE; // 判非法 / mark illegal
END_IF
IF (tStartDelay < T#0S) OR (tStopDelay < T#0S) THEN // 时间窗为负 / a negative time window
    _bCfgBad := TRUE; // 判非法 / mark illegal
END_IF
IF (fFrostLimitC < DL_BHR_FROST_MIN) OR (fFrostLimitC > DL_BHR_FROST_MAX) OR (fFrostLimitC <> fFrostLimitC) THEN // 防霜限温越域 / frost limit out of domain
    _bCfgBad := TRUE; // 判非法 / mark illegal
END_IF
IF (fMinDeltaTC <= 0.0) OR (fMinDeltaTC > DL_BHR_DELTA_MAX) OR (fMinDeltaTC <> fMinDeltaTC) THEN // 最小温差越域 / minimum difference out of domain
    _bCfgBad := TRUE; // 判非法 / mark illegal
END_IF
IF (fEffMinPct < 0.0) OR (fEffMinPct > 100.0) OR (fEffMinPct <> fEffMinPct) THEN // 效率达标阈越域 / efficiency threshold out of domain
    _bCfgBad := TRUE; // 判非法 / mark illegal
END_IF
IF _bCfgBad AND (NOT _bFault) THEN // 组态非法且未锁存 / illegal configuration and not yet latched
    _bFault := TRUE; // 置故障锁存 / raise the fault latch
    _eFaultCause := E_DL_BhrCause.eCfgIllegal; // 故障级成因 (R45 配对 bError) / fault grade cause paired with bError
    _eState := E_DL_BhrState.eFault; // 迁故障相 / migrate to the fault phase
END_IF

// 段 4｜火警联锁：最高优先级，撤命令 + 撤允许 + 锁存 / segment 4, fire alarm interlock with the highest priority
IF bFireAlarm THEN // 火警成立 / the fire alarm is active
    IF NOT _bFault THEN // 未锁存才记故障 / record the fault only when not yet latched
        _bFault := TRUE; // 置故障锁存 / raise the fault latch
        _eFaultCause := E_DL_BhrCause.eFireAlarm; // 故障级成因 (R45 配对 bError) / fault grade cause paired with bError
    END_IF
END_IF

// 段 5｜温度闸与防霜判据：温度非有限即不判防霜（不穿透出口）/ segment 5, temperature gate and frost criterion
_bTempOk := (fExhaustC = fExhaustC) AND ((fExhaustC - fExhaustC) = (fExhaustC - fExhaustC)) AND (fSupplyC = fSupplyC) AND ((fSupplyC - fSupplyC) = (fSupplyC - fSupplyC)) AND (fFreshC = fFreshC) AND ((fFreshC - fFreshC) = (fFreshC - fFreshC)) AND (ABS(fExhaustC) <= DL_BHR_TEMP_MAX) AND (ABS(fFreshC) <= DL_BHR_TEMP_MAX); // 三项温度有限性闸 / finiteness gate on all three temperatures
_bFrost := _bTempOk AND (fFreshC <= fFrostLimitC); // 防霜判据：新风温度低于限温 / frost criterion on the fresh air temperature
_bWheelFbOk := bWheelRunFb AND (NOT bFireAlarm); // 反馈到位判据：反馈有且无火警 / feedback verdict

// 段 6｜相位机：ENUM + CASE，含 ELSE 非法相位兜底（R128）/ segment 6, phase machine with an ELSE fallback for illegal phases
_bConvPermit := FALSE; // 每拍先撤输送允许，只有运行相才能重新置位（防相外残留）/ the permit is withdrawn every scan and only the run phase may raise it again
CASE _eState OF
E_DL_BhrState.eIdle: // 空闲相：有请求且有反馈才进启动等反馈相 / idle, a request plus feedback moves into the start wait
    IF _bFault THEN // 故障锁存 / the fault is latched
        _eState := E_DL_BhrState.eFault; // 迁故障相 / migrate to the fault phase
    ELSIF bConvRunCmd AND bEnable THEN // 有输送请求且使能 / a conveyor request while enabled
        _eState := E_DL_BhrState.eStartWait; // 迁启动等反馈相 / migrate to the start wait phase
    END_IF

E_DL_BhrState.eStartWait: // 启动等反馈相：转轮先启，反馈与延时双满足才放开输送 / start wait, the wheel leads and both feedback and delay must hold
    _bWheelFbOk := bWheelRunFb AND (NOT bFireAlarm) AND _bTempOk; // 本相内反馈判据再收紧（含温度闸）/ the feedback verdict is tightened inside this phase to include the temperature gate
    IF _bFault THEN // 故障锁存 / the fault is latched
        _eState := E_DL_BhrState.eFault; // 迁故障相 / migrate to the fault phase
    ELSIF (NOT bConvRunCmd) THEN // 请求撤销 / the request was withdrawn
        _eState := E_DL_BhrState.eIdle; // 回空闲相 / return to idle
    ELSIF _bWheelFbOk AND tonStart.Q THEN // 反馈到位且启动延时到 / feedback present and the start delay elapsed
        _eState := E_DL_BhrState.eRun; // 迁运行相 / migrate to the run phase
    END_IF

E_DL_BhrState.eRun: // 运行相：输送允许，请求撤销即进吹扫相 / run phase, a withdrawn request moves into purge
    _bConvPermit := bEnable AND bFilterOk AND _bWheelFbOk AND (NOT _bFrost) AND (NOT bFireAlarm); // 输送允许判据，四条判据逐项与 / the conveyor permit is the conjunction of four criteria
    IF _bFault THEN // 故障锁存 / the fault is latched
        _eState := E_DL_BhrState.eFault; // 迁故障相 / migrate to the fault phase
    ELSIF NOT bConvRunCmd THEN // 请求撤销 / the request was withdrawn
        _eState := E_DL_BhrState.ePurge; // 迁吹扫相 / migrate to the purge phase
    END_IF

E_DL_BhrState.ePurge: // 吹扫相：转轮续转，延时到回空闲 / purge phase, the wheel keeps running until the delay elapses
    IF _bFault THEN // 故障锁存 / the fault is latched
        _eState := E_DL_BhrState.eFault; // 迁故障相 / migrate to the fault phase
    ELSIF tonStop.Q THEN // 吹扫延时到 / the purge delay elapsed
        _eState := E_DL_BhrState.eIdle; // 回空闲相 / return to idle
    ELSIF bConvRunCmd THEN // 请求重新给出 / the request is issued again
        _eState := E_DL_BhrState.eStartWait; // 重走启动等反馈相 / restart from the start wait phase
    END_IF

E_DL_BhrState.eFault: // 故障相：全撤命令，等复位沿 / fault phase, all commands withdrawn until the reset edge
    _bConvPermit := FALSE; // 撤输送允许 / the conveyor permit is withdrawn
    _bWheelFbOk := FALSE; // 撤反馈判据 / the feedback verdict is withdrawn

ELSE // 非法相位兜底（R128）/ illegal phase fallback
    _bFault := TRUE; // 置故障锁存 / raise the fault latch
    _eFaultCause := E_DL_BhrCause.eCfgIllegal; // 故障级成因记组态非法 / record the illegal configuration cause
    _eState := E_DL_BhrState.eFault; // 迁故障相 / migrate to the fault phase
    _bConvPermit := FALSE; // 撤输送允许 / the conveyor permit is withdrawn
END_CASE

// 段 7｜转轮命令：启动等反馈 / 运行 / 吹扫三相为真，故障与失能一律撤除 / segment 7, wheel command truth table
bWheelRunCmd := ((_eState = E_DL_BhrState.eStartWait) OR (_eState = E_DL_BhrState.eRun) OR (_eState = E_DL_BhrState.ePurge)) AND bEnable AND (NOT bFireAlarm) AND (NOT _bFault); // 转轮命令，四条件合取 / the wheel command as a conjunction of four conditions
IF _eState = E_DL_BhrState.eFault THEN // 故障相 / the fault phase
    bWheelRunCmd := FALSE; // 撤转轮命令 / withdraw the wheel command
END_IF

// 段 8｜热回收效率：温差不足不更新，出口保持上拍值 / segment 8, heat recovery efficiency with a guarded denominator
IF _bTempOk THEN // 温度可用 / temperatures usable
    _fDeltaT := fExhaustC - fFreshC; // 进排风温差 / the exhaust to fresh difference
    _bEffBaseOk := _fDeltaT >= fMinDeltaTC; // 分母可用判据（含正负方向：仅排风高于新风才有效）/ denominator verdict requiring the exhaust to be warmer than the fresh air
    IF _bEffBaseOk THEN // 分母可用 / the denominator is usable
        _fNum := fSupplyC - fFreshC; // 分子：转轮后温升 / numerator, the temperature rise across the wheel
        _fEff := _fNum / _fDeltaT * 100.0; // 效率，除子已证不小于 fMinDeltaTC / efficiency, divisor proven not below the minimum difference
        IF _fEff < DL_BHR_EFF_MIN THEN // 效率下越界 / efficiency below the floor
            _fEff := DL_BHR_EFF_MIN; // 下钳 / clamp downward
        ELSIF _fEff > DL_BHR_EFF_MAX THEN // 效率上越界 / efficiency above the ceiling
            _fEff := DL_BHR_EFF_MAX; // 上钳 / clamp upward
        END_IF
        IF (_fEff = _fEff) AND ((_fEff - _fEff) = (_fEff - _fEff)) THEN // 结果有限性闸 / result finiteness gate
            _fEffHold := _fEff; // 有效拍更新保持块 / the holder updates on a valid scan
        END_IF
    END_IF
END_IF

// 段 9｜成因分派（固定优先级：故障 > 火警外的降级原因 > 无成因）/ segment 9, cause dispatch with a fixed priority
IF _bFault THEN // 故障锁存优先 / the fault latch takes priority
    eCause := _eFaultCause; // 故障级成因锁存回放 / the fault cause is replayed from the latch
ELSIF _bFrost THEN // 防霜动作 / frost protection tripped
    eCause := E_DL_BhrCause.eFrost; // 信息级成因 / informational cause
ELSIF (NOT bFilterOk) THEN // 过滤网异常 / the filter is unhealthy
    eCause := E_DL_BhrCause.eFilterBad; // 信息级成因 / informational cause
ELSIF (NOT bWheelRunFb) AND (_eState = E_DL_BhrState.eStartWait) THEN // 等反馈相缺反馈 / feedback missing while waiting
    eCause := E_DL_BhrCause.eNoWheelFb; // 信息级成因 / informational cause
ELSIF (NOT _bEffBaseOk) AND _bTempOk THEN // 温差不足 / the temperature difference is too small
    eCause := E_DL_BhrCause.eEffInvalid; // 信息级成因 / informational cause
ELSE
    eCause := E_DL_BhrCause.eNone; // 无成因 / no cause
END_IF

// 段 10｜统一出口 / segment 10, unified outlet
bConvPermit := _bConvPermit AND (_eState = E_DL_BhrState.eRun) AND (NOT _bFault); // 输送允许受运行相与故障锁存双重否决 / the permit is vetoed by the run phase and the fault latch
bFrostProtect := _bFrost; // 防霜动作出口 / frost protection outlet
bWheelFbOk := _bWheelFbOk AND (NOT _bFault); // 反馈到位出口受故障锁存否决 / the feedback outlet is vetoed by the fault latch
fEffPct := _fEffHold; // 效率出口取保持块 / efficiency outlet from the holder
bEffOk := _bEffBaseOk AND (_fEffHold >= fEffMinPct) AND (NOT _bFault); // 效率达标且本拍有效（挂状态量）/ efficiency pass with this scan valid
eState := _eState; // 相位出口单点映射 / single-point phase outlet mapping
bError := _bFault; // 故障标志与锁存位同源 / the fault flag shares the latch source
END_FUNCTION_BLOCK

(* ---- FB_DL_BinderFeederSeq.st ---- *)
(*
  FB_DL_BinderFeederSeq  —  绝缘件振动盘供料顺控（满料/缺料双光电 + 卡料窗） / Binder vibratory feeder sequence with full/empty photoeyes and jam window
  分类 Category : DL_Process
  版本 Version  : 1.0.0
  来源 Source   : t2-2-lbp — 供料/上料工艺族深化
  溯源 Origin   : clean-room 实现，未复制任何源码行
  功能 Function : 1) 三相顺控：eIdle（待机）→ eFeed（供料，bVibOn 输出驱动振动盘，
                  bFullPE 满料到达回 eIdle）→ eFault；使能撤销沿随时回 eIdle；
                  2) 卡料诊断：供料相中缺料（bEmptyPE）持续 tJamWin 未见满料
                  → 0378 卡料锁存（窗为电平式防抖窗，满料到达自动断 IN 复位）；
                  3) 双光电矛盾诊断：bFullPE 与 bEmptyPE 同 TRUE 持续 tContraWin
                  → 0377 矛盾锁存（传感器组态/遮挡异常归因唯一）；
                  4) 信息级三码：供料启动 / 卡料窗激活 / 满料到达（单拍沿）；
                  5) 解除式全当拍量（R240 落地），逐 BOOL 标注见段 4。
  边界 Boundary : ① 组态闸：tJamWin <= 0 或 tContraWin <= 0 → 0376 锁存
                  （组态与 ELSE 兜底归并声明于码表）；
                  ② 满料优先安全侧：矛盾检出期 bVibOn 强制 FALSE（停止振动）；
                  ③ 超时窗均为电平驱动，窗内判据消失自动复位（R176 周期语义合规）；
                  ④ 无 GVL 依赖：纯引脚输入输出，无外部变量引用，无物理 IO 地址。
  依赖 Depends  : Standard.library（TON / R_TRIG）
  码表 Error codes（Process 段 0005，窗口 0376~0378 / 049E~04A0）:
    16#0005_0376 故障级：组态非法（任一窗 <= 0）或相位落 ELSE 兜底（归并声明），锁存至 bReset
    16#0005_0377 故障级：双光电矛盾锁存（满料与缺料同 TRUE 持续 tContraWin），锁存至 bReset
    16#0005_0378 故障级：卡料锁存（供料中缺料持续 tJamWin），锁存至 bReset
    16#0005_049E 信息级：供料启动沿（进 eFeed）
    16#0005_049F 信息级：卡料窗激活沿（供料相缺料进入）
    16#0005_04A0 信息级：满料到达沿（eFeed → eIdle）
  修订历史 Revision :
    2026-11-19  v1.0.0  R42 首版（批次 1 · 序号 3）
*)

TYPE E_DL_BfsState :
(
    eIdle   := 0,    // 待机：满料或未使能 / Idle, full or not enabled
    eFeed   := 10,   // 供料：振动输出驱动 / Feed, vibration output driving
    eFault  := 90    // 故障：卡料或矛盾锁定 / Fault, latched
);
END_TYPE

FUNCTION_BLOCK FB_DL_BinderFeederSeq
VAR_INPUT
    bFeedEn      : BOOL := FALSE;     // 供料使能（电平）[-] / Feed enable, level
    bFullPE      : BOOL := FALSE;     // 满料光电，TRUE = 料满遮挡 [-] / Full photoeye, TRUE = blocked
    bEmptyPE     : BOOL := FALSE;     // 缺料光电，TRUE = 料空遮挡 [-] / Empty photoeye, TRUE = blocked
    tJamWin      : TIME := T#10S;     // 卡料判定窗 [ms]，域 > 0 / Jam detect window
    tContraWin   : TIME := T#500MS;   // 双光电矛盾确认窗 [ms]，域 > 0 / Contradiction confirm window
    bReset       : BOOL := FALSE;     // 复位，上升沿清故障锁存 / Reset edge clears fault latch
END_VAR
VAR_OUTPUT
    eState       : E_DL_BfsState;     // 状态出口，段尾单点映射 / State outlet
    bVibOn       : BOOL;              // 振动盘输出驱动（供料相电平）[-] / Vibrator output drive
    bJamWarn     : BOOL;              // 卡料窗计时中镜像（未到时）[-] / Jam window arming mirror
    bError       : BOOL;              // 故障锁存标志 / Fault latch flag
    nErrId       : UDINT;             // 事件码，0 = 无事件 / Event code
END_VAR
VAR
    tonJam       : TON;               // 卡料判定窗（电平式），无条件刷新 / Jam detect timer
    tonContra    : TON;               // 双光电矛盾确认窗（电平式），无条件刷新 / Contradiction timer
    rtEn         : R_TRIG;            // 使能沿实例，无条件刷新 / Enable edge instance
    rtReset      : R_TRIG;            // 复位沿实例，无条件刷新 / Reset edge instance
    _eState      : E_DL_BfsState := E_DL_BfsState.eIdle;  // 内部相位（CASE 唯一写入目标）/ Internal phase
    _bJamInfoSent: BOOL;              // 卡料窗信息沿单发标志（eFeed 相内保持量）/ Jam-info one-shot sent flag
    _bContra     : BOOL;              // 双光电矛盾当拍量 [-] / Contradiction current-scan flag
    _bFault      : BOOL;              // 故障锁存位（锁存量）/ Latched fault bit
    _uFault      : UDINT;             // 故障码锁存（锁存量）/ Latched fault code
    _uInfo       : UDINT;             // 信息码，每拍重算 / Transient info code
END_VAR

(* —— 段 0：定时器与沿实例无条件周期刷新（禁置于 IF/CASE 内） —— *)
_bContra := bFullPE AND bEmptyPE;                                    // 双光电矛盾（当拍量）
rtEn(CLK := bFeedEn);                                                // 使能沿（每拍必调）
rtReset(CLK := bReset);                                              // 复位沿（每拍必调）
tonJam(IN := (_eState = E_DL_BfsState.eFeed) AND bFeedEn AND bEmptyPE, PT := tJamWin);
                                                // 卡料窗（供料相缺料电平驱动，满料到达自动断 IN）
tonContra(IN := _bContra, PT := tContraWin);
                                                // 矛盾确认窗（矛盾电平驱动，矛盾消失自动断 IN）

(* —— 段 1：单拍量预清零（锁存量 _bFault/_uFault 不入清单，禁同拍抹除） —— *)
_uInfo := 16#0000_0000;             // 信息码每拍重算
bVibOn := FALSE;                    // 振动输出缺省 FALSE（安全侧）
bJamWarn := FALSE;                  // 卡料窗镜像缺省 FALSE
nErrId := 16#0000_0000;             // 事件码缺省无事件

(* —— 段 2：复位沿 + 组态域闸（当拍量判据） —— *)
IF rtReset.Q THEN                   // rtReset.Q = 当拍量
    _bFault := FALSE;               // 清故障锁存位
    _uFault := 16#0000_0000;        // 清故障锁存码
END_IF
IF (TIME_TO_DINT(tJamWin) <= 0) OR (TIME_TO_DINT(tContraWin) <= 0) THEN
    _uFault := 16#0005_0376;        // 故障级：组态非法
    _bFault := TRUE;                // 故障标志与码位配对（R45）
END_IF

(* —— 段 3：矛盾与卡料锁存（判据当拍量/电平式窗） —— *)
IF (NOT _bFault) AND tonContra.Q THEN
    _uFault := 16#0005_0377;        // 故障级：双光电矛盾锁存
    _bFault := TRUE;
END_IF
IF (NOT _bFault) AND tonJam.Q THEN
    _uFault := 16#0005_0378;        // 故障级：卡料锁存
    _bFault := TRUE;
END_IF

(* —— 段 4：故障解除式（R240 落地，逐 BOOL 标注）：
     rtReset.Q = 当拍量；bFeedEn = 当拍量；_bContra = 当拍量；NOT bEmptyPE = 当拍量。
     均不含锁存量（_bFault/_uFault），解除边真实可达：
     矛盾锁存沿「矛盾消失 + 使能撤销 + 复位沿」到达；卡料锁存沿「缺料消失 + 使能撤销 + 复位沿」到达。 —— *)
IF rtReset.Q AND (NOT bFeedEn) AND (NOT _bContra) AND (NOT bEmptyPE) THEN
    _bFault := FALSE;               // 清故障锁存位（锁存量，仅此当拍量解除沿可清）
    _uFault := 16#0000_0000;        // 清故障锁存码（锁存量，仅本当拍量解除沿可清）
    IF _eState = E_DL_BfsState.eFault THEN
        _eState := E_DL_BfsState.eIdle;     // 故障相迁出：回待机
    END_IF
END_IF

(* —— 段 5：相位机（CASE 全覆盖 + ELSE 兜底） —— *)
CASE _eState OF

E_DL_BfsState.eIdle:
    IF rtEn.Q AND (NOT _bFault) AND (NOT _bContra) THEN
        _uInfo := 16#0005_049E;             // 信息级：供料启动沿
        _eState := E_DL_BfsState.eFeed;     // 进供料相
    END_IF

E_DL_BfsState.eFeed:
    bVibOn := bFeedEn AND (NOT _bContra) AND (NOT _bFault);
                                        // 振动输出（矛盾/故障期强制 FALSE，安全侧）
    bJamWarn := bFeedEn AND bEmptyPE AND (NOT tonJam.Q);
                                        // 卡料窗计时中镜像（电平）
    IF bEmptyPE AND (NOT _bJamInfoSent) THEN
        _uInfo := 16#0005_049F;         // 信息级：卡料窗激活沿（单发）
        _bJamInfoSent := TRUE;          // 沿单发标志（eFeed 相内保持）
    END_IF
    IF bFullPE THEN
        _uInfo := 16#0005_04A0;         // 信息级：满料到达沿
        _bJamInfoSent := FALSE;         // 回待机重置单发标志
        _eState := E_DL_BfsState.eIdle; // 满料：回待机相
    ELSIF NOT bFeedEn THEN
        _bJamInfoSent := FALSE;         // 使能撤销：重置单发标志
        _eState := E_DL_BfsState.eIdle; // 回待机相
    END_IF
    (* 卡料/矛盾迁出在段 3 承载 *)

E_DL_BfsState.eFault:
    ;                                   // 故障相：等解除沿（段 4 承载迁出）

ELSE
    _uFault := 16#0005_0376;            // 故障级：非法相位兜底（归并组态码，码表声明）
    _bFault := TRUE;
    _eState := E_DL_BfsState.eFault;    // 强制回故障相

END_CASE

(* —— 段 6：出口单点映射（名实同源；锁存码回放，禁同拍抹除） —— *)
IF _bFault THEN
    nErrId := _uFault;              // 故障锁存码回放
    bVibOn := FALSE;                // 故障相振动输出强制 FALSE（安全侧）
    bJamWarn := FALSE;              // 故障相卡料镜像强制 FALSE（安全侧）
ELSE
    nErrId := _uInfo;               // 信息码
END_IF
bError := _bFault;                  // 故障标志与锁存位同源
eState := _eState;                  // 状态出口单点映射

END_FUNCTION_BLOCK

(* ---- FB_DL_BlindPositionCtrl.st ---- *)
(*==============================================================================
 * 组件名称 (Component)  : FB_DL_BlindPositionCtrl
 * 所属子库 (Sublibrary) : DL_Process
 * 归属目录 (Directory)  : C:\Library\DL_Process
 * 当前版本 (Version)    : 1.0.1
 * 分类/来源标签         : 功能块（FUNCTION_BLOCK）· 暖通遮阳 · 电动帘位置控制
 *                         industry-pool / hvac / shading / interlock
 * 兼容性   (Platform)   : CODESYS 3.5 / TwinCAT 3 / 汇川 InoProShop / 施耐德
 *                         Machine Expert；仅用 Standard.library 的 TON
 * 溯源声明 (Provenance) : 道莅自研 clean-room——只借公开规范条款与工程惯例，零代码行复制。
 * 【R33 已返修】安全相方向 / 位置记账 / 到位判据三者同向：eSafeRetract 改驱动
 *                         上行（oMotorUp），与位置递减记账、bUpLimitSw 到位判据一致。
 * 功能一句话 (Summary)  : 电动遮阳帘位置控制：位置指令按行程时间标定估计，
 *                         风雨联锁强制收回到底，结冰联锁冻结驱动，限位开关校准。
 *
 * 功能描述 (Function)   : 五态状态机：空闲/上行/下行/保持/安全收回。位置估计
 *                         用 100ms 节拍累计行程时间比例（每拍加 100ms/全程
 *                         时间 × 100），限位开关到位即校准端点；风雨联锁任一
 *                         为真立即转安全收回（驱动上行至下限位全收）；结冰联锁
 *                         冻结驱动输出并报故障；行程时间域外标定无效报故障。
 * 与既有件边界 (Boundary): 借 OSCAT BLIND 的行为定义（光照目标 + 风雨联锁 +
 *                         行程时间标定），clean-room 实现；光照闭环采样归
 *                         上层调度，本件只接位置指令。
 * 码位说明 (Codes)      : 信息 16#0006_300F 安全收回激活（风雨联锁）
 *                         故障 16#0006_3010 行程时间域外，标定无效
 *                         故障 16#0006_3011 输出互锁校验失败（上下同出）
 *                         故障 16#0006_3012 结冰联锁，驱动已冻结
 *                         段 16#06_0_0F~13 首槽信息级、次槽起故障级。
 * 依赖说明 (Depends)    : 无 DL_ 内部依赖；仅 Standard.library 的 TON / ABS。
 * 红线自检 (Redline)    : 零全局依赖 ｜ 零 VAR_EXTERNAL ｜ 零 %I/%Q（输出引脚）
 *                         浮点比较带 fEps 容差 ｜ ENUM 配 CASE 且 ELSE 兜底
 *                         定时器每周期无条件刷新 ｜ 全变量双语同行注释
 *                         安全联锁（风雨冰）在 CASE 之前最高优先拦截
 * 修订历史 (Revision)   : 2026-11-18  v1.0.0  首版入库（R32 · 批 3）
 *                        2026-11-18  v1.0.1  R33 返修：安全相驱动方向与记账/到位判据同向、节拍计时自复位
 *============================================================================*)

FUNCTION_BLOCK FB_DL_BlindPositionCtrl
VAR_INPUT
    bRun         : BOOL;                    // 控制使能，假则停驱动回空闲 / Enable, FALSE stops and idles
    iCmdPosPct   : INT;                     // 位置指令 [％]，域 0 到 100，0 全收 100 全开 / Position command, 0 to 100
    bWindAlarm   : BOOL;                    // 风速联锁 [事件]，真则强制收回 / Wind interlock, TRUE forces retract
    bRainAlarm   : BOOL;                    // 雨水联锁 [事件]，真则强制收回 / Rain interlock, TRUE forces retract
    bIceAlarm    : BOOL;                    // 结冰联锁 [事件]，真则冻结驱动 / Ice interlock, TRUE freezes the drive
    bUpLimitSw   : BOOL;                    // 上限位开关 [开关]，真为全收到位 / Upper limit switch, fully retracted
    bDnLimitSw   : BOOL;                    // 下限位开关 [开关]，真为全开到位 / Lower limit switch, fully extended
    fTravelTimeS : LREAL := 60.0;           // 全程运行时间 [s]，标定参数 / Full travel time, calibration
    fEps         : LREAL := 1.0E-6;         // 浮点判零容差 [实数域] / Floating zero tolerance
END_VAR
VAR_OUTPUT
    oMotorUp : BOOL;                    // 电机上行输出 [引脚]，经适配层映射 / Motor up output
    oMotorDn : BOOL;                    // 电机下行输出 [引脚]，经适配层映射 / Motor down output
    iEstPosPct: INT;                    // 估计位置 [％]，行程时间标定 / Estimated position
    eState   : (eIdle := 0, eMovingUp := 1, eMovingDown := 2, eHoldPos := 3, eSafeRetract := 4);  // 状态枚举输出 / State output
    bError   : BOOL;                    // 故障标志，与故障码配对 / Fault flag paired with codes
    uErrorId : UDINT;                   // 事件码，0 表示无事件 / Event code, zero means none
END_VAR
VAR
    tonPace  : TON;     // 行程估计节拍定时器 [s]，每拍无条件刷新 / Travel pace timer
    fStepPct : LREAL;   // 单节拍位置步进 [％] / Position step per pace tick
    iPosF    : LREAL;   // 估计位置浮点内部值 [％] / Estimated position, internal float
    bCalOk   : BOOL;    // 行程标定有效标志 / Calibration validity flag
    uCodeLatch: UDINT;  // 故障锁存码 [码] / Latched fault code
    uInfoCode: UDINT;   // 信息级单拍码 [码] / One-shot info code
END_VAR
VAR CONSTANT
    DL_BPC_PACE_MS : TIME := T#100MS;   // 行程估计节拍 [ms] / Travel pace period
    DL_BPC_PACES   : LREAL := 0.1;      // 节拍秒值 [s]，与 PACE_MS 一致 / Pace in seconds
    DL_BPC_MAXTT   : LREAL := 3600.0;   // 行程时间上限 [s]，防标定离谱 / Travel time cap
END_VAR

(* 段 1｜定时器无条件刷新与标定域闸（红线 7）/ Timer refresh and calibration gate *)
tonPace(IN := NOT tonPace.Q, PT := DL_BPC_PACE_MS);     // 节拍自复位振荡（红线 7）/ Self-reset oscillating pace
IF (fTravelTimeS > fEps) AND (fTravelTimeS <= DL_BPC_MAXTT) THEN
    bCalOk := TRUE;                 // 标定有效 / Calibration valid
    fStepPct := DL_BPC_PACES / fTravelTimeS * 100.0;    // 单拍步进导出 / Step per tick
ELSE
    bCalOk := FALSE;                // 标定无效 / Calibration invalid
    fStepPct := 0.0;                // 步进置零禁走 / Zero step, no motion
    uCodeLatch := 16#0006_3010;     // 故障级：标定无效 / Fault: invalid calibration
END_IF

(* 段 2｜最高优先级安全联锁（先于 CASE）：风雨强收、结冰冻结 / Highest-priority safety before the CASE *)
IF bIceAlarm THEN
    oMotorUp := FALSE;              // 冻结上行 / Freeze up
    oMotorDn := FALSE;              // 冻结下行 / Freeze down
    IF bCalOk THEN
        uCodeLatch := 16#0006_3012; // 故障级：结冰冻结（标定有效才报）/ Fault: ice freeze
    END_IF
    eState := eHoldPos;             // 拍 N 保持位置，拍 N+1 由 CASE 复核 / Hold this scan
ELSIF bWindAlarm OR bRainAlarm THEN
    uInfoCode := 16#0006_300F;      // 信息级：安全收回激活 / Info: safe retract active
    eState := eSafeRetract;         // 拍 N 转安全收回，拍 N+1 执行 / To safe retract
END_IF

(* 段 3｜状态机主分派（ENUM 配 CASE，ELSE 兜底）/ State dispatch with ELSE interception *)
CASE eState OF

    eIdle:
        (* 本拍行为：停驱动；指令与使能俱备且不在联锁期拍 N+1 起步 / Stop; start when commanded *)
        oMotorUp := FALSE;              // 停上行 / Stop up
        oMotorDn := FALSE;              // 停下行 / Stop down
        IF bRun AND bCalOk AND (NOT bIceAlarm) AND (NOT bWindAlarm) AND (NOT bRainAlarm) THEN
            IF (iCmdPosPct > iEstPosPct) AND (iCmdPosPct <= 100) THEN
                eState := eMovingDown;  // 指令更大：向全开方向 / Bigger command: extend
            ELSIF (iCmdPosPct < iEstPosPct) AND (iCmdPosPct >= 0) THEN
                eState := eMovingUp;    // 指令更小：向全收方向 / Smaller command: retract
            ELSE
                eState := eHoldPos;     // 已在目标位保持 / Hold at target
            END_IF
        END_IF

    eMovingUp:
        (* 本拍行为：驱动上行并累计位置；到位或到目标转保持 / Drive up and accumulate; stop at target *)
        IF NOT (bRun AND bCalOk) THEN
            eState := eIdle;            // 撤使能或标定失效回空闲 / Disable or bad calibration to idle
        ELSE
            oMotorUp := TRUE;           // 驱动上行 / Drive up
            oMotorDn := FALSE;          // 下行必停 / Down must be off
            IF tonPace.Q THEN
                iPosF := iPosF - fStepPct;      // 位置递减（上行） / Position decreases
            END_IF
            IF bUpLimitSw OR (iPosF <= 0.0) THEN
                iPosF := 0.0;           // 全收校准端点 / Calibrate the endpoint
                oMotorUp := FALSE;      // 停驱动 / Stop the drive
                eState := eHoldPos;     // 拍 N+1 保持 / Hold next scan
            ELSIF iPosF <= DINT_TO_LREAL(iCmdPosPct) THEN
                oMotorUp := FALSE;      // 到目标停 / Stop at the target
                eState := eHoldPos;
            END_IF
        END_IF

    eMovingDown:
        (* 本拍行为：驱动下行并累计位置；到位或到目标转保持 / Drive down and accumulate *)
        IF NOT (bRun AND bCalOk) THEN
            eState := eIdle;            // 撤使能回空闲 / Disable to idle
        ELSE
            oMotorUp := FALSE;          // 上行必停 / Up must be off
            oMotorDn := TRUE;           // 驱动下行 / Drive down
            IF tonPace.Q THEN
                iPosF := iPosF + fStepPct;      // 位置递增（下行）/ Position increases
            END_IF
            IF bDnLimitSw OR (iPosF >= 100.0) THEN
                iPosF := 100.0;         // 全开校准端点 / Calibrate the endpoint
                oMotorDn := FALSE;      // 停驱动 / Stop the drive
                eState := eHoldPos;     // 拍 N+1 保持 / Hold next scan
            ELSIF iPosF >= DINT_TO_LREAL(iCmdPosPct) THEN
                oMotorDn := FALSE;      // 到目标停 / Stop at the target
                eState := eHoldPos;
            END_IF
        END_IF

    eHoldPos:
        (* 本拍行为：停驱动监视指令；新指令转移动相 / Hold and watch the command *)
        oMotorUp := FALSE;              // 停上行 / Stop up
        oMotorDn := FALSE;              // 停下行 / Stop down
        IF bRun AND bCalOk AND (NOT bIceAlarm) AND (NOT bWindAlarm) AND (NOT bRainAlarm) THEN
            IF (iCmdPosPct > iEstPosPct) AND (iCmdPosPct <= 100) THEN
                eState := eMovingDown;  // 起步向全开 / Start to extend
            ELSIF (iCmdPosPct < iEstPosPct) AND (iCmdPosPct >= 0) THEN
                eState := eMovingUp;    // 起步向全收 / Start to retract
            END_IF
        END_IF

    eSafeRetract:
        (* 本拍行为：驱动上行收回到底（与位置递减记账、bUpLimitSw 到位判据同向）；联锁撤清且到位转保持
         * Drive up to fully retracted, same direction as the decreasing position bookkeeping and bUpLimitSw *)
        oMotorDn := FALSE;              // 下行必停 / Down must be off
        oMotorUp := TRUE;               // 强制上行收回（与记账递减同向）/ Forced up retract, same direction
        IF tonPace.Q THEN
            iPosF := iPosF - fStepPct;  // 收回位置递减 / Retract position decreases
        END_IF
        IF bUpLimitSw OR (iPosF <= 0.0) THEN
            iPosF := 0.0;               // 全收校准 / Calibrate fully retracted
            oMotorUp := FALSE;          // 停驱动 / Stop the drive
            eState := eHoldPos;         // 拍 N+1 保持 / Hold next scan
        END_IF

ELSE
    oMotorUp := FALSE;                  // 非法状态双输出必停 / Illegal state, both off
    oMotorDn := FALSE;
    eState := eIdle;                    // 拦截回空闲 / Intercept to idle
    uCodeLatch := 16#0006_3010;         // 故障：状态越界 / Fault: state out of range
END_CASE

(* 段 4｜输出互锁校验（防御闸）与出口装配 / Interlock check and exit assembly *)
IF oMotorUp AND oMotorDn THEN
    oMotorUp := FALSE;                  // 互锁失败双断 / Interlock failure, both off
    oMotorDn := FALSE;
    uCodeLatch := 16#0006_3011;         // 故障级：互锁校验失败 / Fault: interlock broken
END_IF
iEstPosPct := LREAL_TO_DINT(iPosF);     // 估计位置整数输出 / Integer position output
IF iEstPosPct < 0 THEN
    iEstPosPct := 0;                    // 钳下界 / Clamp low
ELSIF iEstPosPct > 100 THEN
    iEstPosPct := 100;                  // 钳上界 / Clamp high
END_IF
IF NOT bRun THEN
    uCodeLatch := 16#0000_0000;         // 撤使能清标定故障（可达解除）/ Run drop clears faults
END_IF
bError := (uCodeLatch <> 16#0000_0000); // 故障锁存回放 / Latched fault replay
IF uCodeLatch <> 16#0000_0000 THEN
    uErrorId := uCodeLatch;             // 故障码优先 / Fault first
    uInfoCode := 16#0000_0000;
ELSE
    uErrorId := uInfoCode;              // 信息码单拍 / Info one shot
    uInfoCode := 16#0000_0000;
END_IF
END_FUNCTION_BLOCK

(* ---- FB_DL_BoilerBlowdownSeq.st ---- *)
(*==============================================================================
 * 组件名称 (Component)  : FB_DL_BoilerBlowdownSeq
 * 所属子库 (Sublibrary) : DL_Process
 * 当前版本 (Version)    : 1.0.0
 * 兼容性   (Platform)   : CODESYS 3.5+ / TwinCAT 3 / 汇川 InoProShop / 施耐德 Machine Expert
 *                         仅依赖 Standard.library（TON / R_TRIG / ABS），零厂商私有库
 * 功能描述 (Function)   : 锅炉排污顺控。触发源三选一：定时（tInterval 到）／电导率超
 *                         fCondLimitUs／手动 bManTrigger 上升沿 → eOpen（开排污阀，时长 tBlowTime，
 *                         单次硬上限 tBlowMax）→ eSettle（关阀后稳定 tSettleTime）→ eDone。
 *                         联锁：低水位 bLevelLow 为真 → **禁止开启**（干烧风险）；若排污中水位转低
 *                         则立即关阀并置故障；排污期间水位下降量超 fLevelDropMaxPct → 中止并置码。
 * 接口     (Interface)  : 输入 bEnable 使能、tInterval 定时排污周期、fCondUs 实测电导率、
 *                         fCondLimitUs 电导率上限、bManTrigger 手动触发、bLevelLow 低水位联锁、
 *                         fLevelPct 水位、fLevelDropMaxPct 排污期允许水位降幅、tBlowTime 排污时长、
 *                         tBlowMax 单次排污硬上限、tSettleTime 关阀稳定时长、bReset 复位；
 *                         输出 bValveCmd 排污阀命令、nBlowCount 累计排污次数（锁存量，复位不清零）、
 *                         eState、eCause、bError、nErrId。
 * 边界     (Boundary)   : ① 组态闸：tBlowTime <= T#0S、tBlowMax <= tBlowTime、tInterval <= T#0S、
 *                         fCondLimitUs <= 0.0、fLevelDropMaxPct <= 0.0、tSettleTime <= T#0S 或任一
 *                         浮点引脚 NaN → 故障锁存，**且非法时 bValveCmd 直接为 FALSE**（安全侧：阀关）；
 *                         ② 排污水量/时长硬钳位：单次 PT = MIN(tBlowTime, tBlowMax)，防卡阀长时间
 *                         排污把锅炉抽空（钳在 PT 而非事后判，结构性杜绝超时溢流）；
 *                         ③ **周期定时器自复位**：tonInterval 的 IN := NOT tonInterval.Q（R188），
 *                         不依赖外部沿清零，节拍窗永不卡死；
 *                         ④ TON 三枚 + R_TRIG 三枚段 0 无条件周期刷新（R228A）；
 *                         ⑤ 故障相迁出唯一路径 = bReset 上升沿；⑥ 零全局耦合（无 GVL / 无物理地址）。
 * 解除式   (Release)    : bReset 上升沿 ∧ 组态合法 ∧ 水位已恢复（bLevelLow = FALSE 且水位降幅
 *                         已回落到 fLevelDropMaxPct 之内，均为当拍量，R240 范式）。
 *                         自证可满足（终审两式 1）：三枚 TON 的 IN 挂相位，故障相内恒假 → Q 恒假；
 *                         水位回升由补水泵保证（外部职责），故路径物理可达、无恒假因子。
 * 码表     (Codes)      : 16#0005_03A8 故障级：排污顺控故障总码（组态非法 / 低水位联锁 /
 *                         水位降幅超限 / 非法相位），锁存至 bReset 上升沿，归因由 eCause 承载
 *                         （R190 单件单总码，各成因独立赋值点）；16#0005_04D0 信息级：单次排污完成。
 *                         加码反证（R90）：完成时 bValveCmd 已关、eState 驻留 eDone，与「一直待在
 *                         eDone」出口同值；累计次数 nBlowCount 的变化虽可观测，但它是累计台账，
 *                         无法分辨当前这一次归零，故立一码记录每次排污动作的完成沿。
 *                         码段说明：0005 段故障子带 03xx / 信息子带 04xx，本件取 03A8 / 04D0
 *                         （源码实扫该两槽为空，续接同子带已用最大值，未回填碎片孔洞）。
 * 开源溯源 (Origin)     : 道莅自研 clean-room（参考锅炉排污公用工程语义与参数域，
 *                         零代码行复制；t1-2-oscat-building 族）
 * 修订历史 (Revision)   : 2026-11-19  v1.0.0  R45 首版（批次 4 · 序号 20）
 *==============================================================================*)

TYPE E_DL_BbsState :
(
    eIdle   := 0,     // 待触发（阀关） / Idle, valve closed
    eOpen   := 10,    // 排污阀开启计时 / Blowdown valve open
    eSettle := 20,    // 关阀后稳定 / Settling after valve closure
    eDone   := 30,    // 本次排污完成 / Blowdown done
    eFault  := 90     // 故障锁存相（阀关） / Fault latched phase, valve closed
);
END_TYPE

TYPE E_DL_BbsCause :
(
    eNone         := 0,  // 无故障成因 / No cause
    eCfgIllegal   := 1,  // 组态非法 / Illegal configuration
    eLevelLowLock := 2,  // 低水位联锁（禁止开启或中途关阀） / Low-level interlock
    eLevelDrop    := 3,  // 排污期水位降幅超限 / Level drop over limit during blowdown
    ePhaseBad     := 4   // 非法相位兜底 / Illegal phase fallback
);
END_TYPE

FUNCTION_BLOCK FB_DL_BoilerBlowdownSeq
VAR_INPUT
    bEnable         : BOOL := TRUE;       // 排污功能使能 [-] / Blowdown enabled
    tInterval       : TIME := T#8H;       // 定时排污周期，域 > T#0S [ms] / Periodic blowdown interval [ms]
    fCondUs         : REAL := 0.0;        // 实测电导率 [µS/cm] / Measured conductivity [uS/cm]
    fCondLimitUs    : REAL := 3000.0;     // 电导率上限（超限触发排污），域 > 0.0 [µS/cm] / Conductivity limit, domain > 0.0 [uS/cm]
    bManTrigger     : BOOL := FALSE;      // 手动触发（上升沿有效） [-] / Manual trigger, rising edge
    bLevelLow       : BOOL := FALSE;      // 低水位联锁（TRUE 禁止开启，已开立即关阀） [-] / Low-level interlock
    fLevelPct       : REAL := 60.0;       // 水位 [%] / Water level [%]
    fLevelDropMaxPct: REAL := 8.0;        // 排污期允许水位降幅，域 > 0.0 [%] / Allowed level drop during blowdown [%]
    tBlowTime       : TIME := T#30S;      // 单次排污时长，域 > T#0S [ms] / Blowdown duration [ms]
    tBlowMax        : TIME := T#60S;      // 单次排污硬上限，域 > tBlowTime [ms] / Hard blowdown ceiling [ms]
    tSettleTime     : TIME := T#10S;      // 关阀稳定时长，域 > T#0S [ms] / Post-close settling time [ms]
    bReset          : BOOL := FALSE;      // 复位命令，上升沿清故障（不清累计次数） [-] / Reset clears fault, count preserved
END_VAR
VAR_OUTPUT
    bValveCmd       : BOOL;               // 排污阀命令（故障/组态非法恒 FALSE） [-] / Blowdown valve command, FALSE in fault
    nBlowCount      : UDINT;              // 累计排污次数（锁存量，复位不清零） [次] / Cumulative blowdown count, kept across resets
    eState          : E_DL_BbsState;      // 状态出口，段 6 单点映射 / State outlet
    eCause          : E_DL_BbsCause;      // 故障成因出口（R190 归因唯一） / Fault cause outlet
    bError          : BOOL;               // 故障锁存标志 [-] / Fault latch flag
    nErrId          : UDINT;              // 事件码，0 = 无事件 / Event code, 0 = no event
END_VAR
VAR
    _eState         : E_DL_BbsState := E_DL_BbsState.eIdle;   // 内部相位（CASE 唯一写入目标） / Internal phase
    _eCause         : E_DL_BbsCause := E_DL_BbsCause.eNone;   // 故障成因锁存（锁存量） / Latched cause
    tonInterval     : TON;                // 周期定时（自复位），段 0 无条件调用 / Self-resetting interval timer
    tonBlow         : TON;                // 排污计时（PT 已硬钳位），段 0 无条件调用 / Blowdown timer with clamped preset
    tonSettle       : TON;                // 关阀稳定计时，段 0 无条件调用 / Settle timer
    rtMan           : R_TRIG;             // 手动触发沿实例，段 0 无条件调用 / Manual trigger edge
    rtLevelLow      : R_TRIG;             // 低水位上升沿实例，段 0 无条件调用 / Low-level rising edge
    rtReset         : R_TRIG;             // 复位沿实例，段 0 无条件调用 / Reset edge
    _tBlowPreset    : TIME;               // 排污计时预置（MIN(tBlowTime, tBlowMax) 当拍量） [ms] / Clamped blowdown preset [ms]
    _fLevelAtStart  : REAL;               // 排污起始水位快照（锁存量） [%] / Level snapshot at blowdown start, latched
    _bSnapshotOk    : BOOL;               // 起始水位快照有效（锁存量） [-] / Start-level snapshot valid
    _fLevelDrop     : REAL;               // 本次水位降幅（当拍量） [%] / Level drop this blowdown [%]
    _nBlowCount     : UDINT;              // 累计排污次数（锁存量，复位不清零） [次] / Cumulative count, kept across resets
    _bCondOver      : BOOL;               // 电导率超限当拍量 [-] / Conductivity over limit
    _bNonFin        : BOOL;               // 输入非有限当拍量 [-] / Non-finite input this scan
    _bCfgBad        : BOOL;               // 组态非法当拍量 [-] / Illegal configuration
    _bDropExcess    : BOOL;               // 水位降幅超限当拍量 [-] / Level drop over limit
    _bLevelOk       : BOOL;               // 水位已恢复当拍量（解除可达性判据） [-] / Level recovered verdict
    _bFault         : BOOL;               // 故障锁存位（锁存量） / Latched fault bit
    _uFault         : UDINT;              // 故障码锁存（锁存量） / Latched fault code
    _uInfo          : UDINT;              // 信息码，每拍重算 / Info code, recomputed each scan
END_VAR
VAR CONSTANT
    DL_COUNT_MAX : UDINT := 16#FFFF_FFFE; // 累计次数饱和上限，留加 1 裕度防溢出 [次] / Count saturation limit with margin [count]
END_VAR

(* —— 段 0：当拍判据派生 + 3 枚 TON（含自复位周期定时）与 3 枚 R_TRIG 无条件刷新 —— *)
IF tBlowTime < tBlowMax THEN                                             // 硬钳位：取小者，结构性防超时溢流 / Hard clamp to the smaller preset
    _tBlowPreset := tBlowTime;
ELSE
    _tBlowPreset := tBlowMax;
END_IF
_bCondOver := fCondUs > fCondLimitUs;                                    // 电导率超限当拍量 / Conductivity over limit
_bNonFin   := (fCondUs <> fCondUs) OR (fLevelPct <> fLevelPct)           // NaN 自反判（判等禁令唯一例外） / NaN self-reflexive tests
           OR (fCondLimitUs <> fCondLimitUs) OR (fLevelDropMaxPct <> fLevelDropMaxPct);
_fLevelDrop := _fLevelAtStart - fLevelPct;                               // 本次水位降幅 / Level drop this blowdown
_bDropExcess := _bSnapshotOk AND (_fLevelDrop > fLevelDropMaxPct);       // 降幅超限当拍量 / Drop over limit
_bLevelOk := (NOT bLevelLow) AND ((NOT _bSnapshotOk) OR (_fLevelDrop <= fLevelDropMaxPct));   // 水位已恢复（解除判据） / Level recovered
_bCfgBad := (tBlowTime <= T#0S) OR (tBlowMax <= tBlowTime) OR (tInterval <= T#0S)              // 时间正域与配比闸（R151） / Time gates and ratio constraints
            OR (fCondLimitUs <= 0.0) OR (fLevelDropMaxPct <= 0.0) OR (tSettleTime <= T#0S);     // 浮点与稳定时间闸 / Float and settle gates
rtMan(CLK := bManTrigger);                                                                     // 手动沿，每拍必调（R228A） / Manual edge
rtLevelLow(CLK := bLevelLow);                                                                   // 低水位沿，每拍必调 / Low-level edge
rtReset(CLK := bReset);                                                                         // 复位沿，每拍必调 / Reset edge
tonInterval(IN := NOT tonInterval.Q, PT := tInterval);                                          // 周期定时自复位（R188），IN 取自身 Q 反 / Self-resetting interval timer
tonBlow(IN := (_eState = E_DL_BbsState.eOpen), PT := _tBlowPreset);                             // 排污计时（PT 已钳位，IN 绑相位） / Blowdown timer
tonSettle(IN := (_eState = E_DL_BbsState.eSettle), PT := tSettleTime);                          // 关阀稳定计时（IN 绑相位） / Settle timer

(* —— 段 1：单拍量预清零（锁存量不入清单，R107） —— *)
_uInfo       := 16#0000_0000;      // 信息码每拍重算 / Info recomputed every scan
bValveCmd    := FALSE;             // 阀命令缺省关（安全侧，任何分支须显式开） / Valve defaults closed, safe side
nBlowCount   := _nBlowCount;       // 累计次数镜像（锁存量回放，复位不清零） / Cumulative count mirror
nErrId       := 16#0000_0000;      // 事件码缺省无事件 / Event code default none
bError       := FALSE;             // 故障标志每拍预清，故障分支同拍置位（R45 配对） / Flag preset

(* —— 段 2：复位沿 + 组态域闸 + 低水位联锁 —— *)
IF rtReset.Q THEN                                                        // 当拍复位沿 / current-scan reset edge
    _bFault := FALSE;                                                    // 清故障锁存位（锁存量） / Clear fault latch
    _uFault := 16#0000_0000;                                             // 清故障锁存码（锁存量） / Clear latched code
    _eCause := E_DL_BbsCause.eNone;                                      // 清成因（锁存量） / Clear latched cause
    _bSnapshotOk := FALSE;                                               // 起始水位快照重新武装 / Re-arm the start-level snapshot
    IF _eState = E_DL_BbsState.eFault THEN
        _eState := E_DL_BbsState.eIdle;                                  // 故障相迁出唯一路径 / Sole exit from fault phase
    END_IF
END_IF
IF _bCfgBad OR _bNonFin THEN                                             // 组态非法（含非有限） → 故障且阀关 / Illegal config, fault with valve closed
    _uFault := 16#0005_03A8;                                             // 故障级：排污顺控故障总码 / Fault-level: blowdown fault code
    _bFault := TRUE;
    bError  := TRUE;                                                     // 故障标志同拍置位（R45 配对） / Error flag set same scan
    _eCause := E_DL_BbsCause.eCfgIllegal;                                // 归因：组态非法 / Cause: illegal configuration
END_IF
IF (NOT _bFault) AND bLevelLow THEN                                      // 低水位联锁：禁止开启；已开则立即关阀 / Low-level interlock
    _uFault := 16#0005_03A8;
    _bFault := TRUE;
    bError  := TRUE;
    _eCause := E_DL_BbsCause.eLevelLowLock;                              // 归因：低水位联锁 / Cause: low-level interlock
END_IF
IF (NOT _bFault) AND _bDropExcess THEN                                   // 排污期水位降幅超限 → 中止 / Level drop over limit, abort
    _uFault := 16#0005_03A8;
    _bFault := TRUE;
    bError  := TRUE;
    _eCause := E_DL_BbsCause.eLevelDrop;                                 // 归因：水位降幅超限 / Cause: level drop over limit
END_IF

(* —— 段 3：故障解除式（R240 全当拍量） —— *)
IF rtReset.Q AND (NOT _bCfgBad) AND (NOT _bNonFin) AND _bLevelOk THEN
    _bFault := FALSE;                                                    // 清故障锁存位（锁存量） / Clear fault latch
    _uFault := 16#0000_0000;                                             // 清故障锁存码（锁存量） / Clear latched code
    _eCause := E_DL_BbsCause.eNone;                                      // 清成因（锁存量） / Clear latched cause
END_IF

(* —— 段 3A：故障锁存相位迁移闸 —— *)
IF _bFault AND (_eState <> E_DL_BbsState.eFault) THEN
    _eState := E_DL_BbsState.eFault;                                     // 锁存即入故障相 / Latch enters fault phase
END_IF

(* —— 段 4：相位机（ENUM 全成员显式标签 + ELSE 兜底，R128） —— *)
CASE _eState OF

E_DL_BbsState.eIdle:
    IF (NOT bEnable) THEN                                                // 出口 1：未使能，明确驻留 / Disabled, explicit stay
        _eState := E_DL_BbsState.eIdle;
    ELSIF (NOT _bFault) AND (NOT bLevelLow)                              // 出口 2：三触发源之一命中且水位允许 / Any of the three triggers with level permission
          AND (tonInterval.Q OR _bCondOver OR rtMan.Q) THEN
        (* 周期窗无需手动复位：tonInterval 的 IN := NOT Q 自复位，下一拍自动重走一窗（R188） / The interval window self-restarts, no manual reset *)
        _fLevelAtStart := fLevelPct;                                     // 锁存起始水位（唯一写入点） / Latch the start level
        _bSnapshotOk := TRUE;                                            // 快照有效 / Snapshot valid
        _eState := E_DL_BbsState.eOpen;                                  // 进排污相 / Enter blowdown phase
    ELSIF _bFault THEN                                                   // 出口 3：故障锁存 / Fault latched
        _eState := E_DL_BbsState.eFault;
    END_IF

E_DL_BbsState.eOpen:
    IF tonBlow.Q THEN                                                    // 出口 1：排污时长到 / Blowdown time elapsed
        _eState := E_DL_BbsState.eSettle;
    ELSIF bLevelLow THEN                                                 // 出口 2：水位转低（前置消失，R98；故障由段 2 置） / Level low during blowdown
        _eState := E_DL_BbsState.eFault;
    END_IF

E_DL_BbsState.eSettle:
    IF tonSettle.Q THEN                                                  // 出口 1：稳定时长到 / Settle time elapsed
        IF _nBlowCount < DL_COUNT_MAX THEN
            _nBlowCount := _nBlowCount + 1;                              // 累计排污次数递增（单点写入） / Cumulative count increment
        END_IF
        _uInfo := 16#0005_04D0;                                          // 信息级：单次排污完成 / Info: one blowdown completed
        _eState := E_DL_BbsState.eDone;
    ELSIF bLevelLow THEN                                                 // 出口 2：稳定期水位转低 / Level low while settling
        _eState := E_DL_BbsState.eIdle;
    END_IF

E_DL_BbsState.eDone:
    IF (NOT bEnable) OR bLevelLow THEN                                   // 出口 1：未使能或水位低，回空闲 / Disabled or level low returns idle
        _eState := E_DL_BbsState.eIdle;
    ELSIF _bFault THEN                                                   // 出口 2：故障锁存 / Fault latched
        _eState := E_DL_BbsState.eFault;
    END_IF

E_DL_BbsState.eFault:
    ;                                                                     // 故障相：仅段 3 复位沿可迁出 / Only the reset edge leaves this phase

ELSE
    _uFault := 16#0005_03A8;                                             // 故障级：非法相位兜底（归并总码） / Illegal-phase fallback
    _bFault := TRUE;
    bError  := TRUE;
    _eCause := E_DL_BbsCause.ePhaseBad;                                  // 归因：非法相位 / Cause: illegal phase
    _eState := E_DL_BbsState.eFault;

END_CASE

(* —— 段 5：出口单点映射（名实同源；锁存码回放；阀安全侧） —— *)
IF _bFault OR _bCfgBad OR (NOT bEnable) OR bLevelLow THEN
    bValveCmd := FALSE;                                                  // 故障/组态非法/失能/低水位：阀恒关 / Valve forced closed
ELSE
    bValveCmd := (_eState = E_DL_BbsState.eOpen);                        // 仅排污相开阀 / Valve open only in the blowdown phase
END_IF
IF _bFault THEN
    nErrId := _uFault;                                                   // 故障锁存码回放 / Replay latched fault code
ELSE
    nErrId := _uInfo;                                                    // 信息码 / Info code
END_IF
bError := _bFault;                                                       // 故障标志与锁存同源（名实双出口，R191） / Flag from latch
eState := _eState;                                                       // 状态出口 / State outlet
eCause := _eCause;                                                       // 成因出口 / Cause outlet

END_FUNCTION_BLOCK
